(* IEC 61131-3 sources: plc-st-coding-agent/progress/evidence/f14_v3_parallel_20261112/jobs/custom_deepseek-v4pro, 102 files *)

(* ---- public-easy-01.candidate_01.st ---- *)
FUNCTION_BLOCK AutomatedFillingLineControl
VAR_INPUT
    bottleSensor : BOOL;
    cleaningConfirmButton : BOOL;
    fillingConfirmButton : BOOL;
    cappingConfirmButton : BOOL;
    packingConfirmButton : BOOL;
    finishedButton : BOOL;
END_VAR
VAR_OUTPUT
    Pump_Motor : BOOL;
    Filling_Valve : BOOL;
    Capping_Machine : BOOL;
    Packing_Machine : BOOL;
    Completion_Light : BOOL;
END_VAR
VAR
    state : INT := 0; (* 0=Idle, 1=Cleaning, 2=Filling, 3=Capping, 4=Packing, 5=Completed *)
END_VAR

CASE state OF
    0: (* Idle *)
        Pump_Motor := FALSE;
        Filling_Valve := FALSE;
        Capping_Machine := FALSE;
        Packing_Machine := FALSE;
        Completion_Light := FALSE;
        IF bottleSensor THEN
            state := 1;
        END_IF;

    1: (* Cleaning *)
        Pump_Motor := TRUE;
        Filling_Valve := FALSE;
        Capping_Machine := FALSE;
        Packing_Machine := FALSE;
        Completion_Light := FALSE;
        IF cleaningConfirmButton THEN
            state := 2;
        END_IF;

    2: (* Filling *)
        Pump_Motor := FALSE;
        Filling_Valve := TRUE;
        Capping_Machine := FALSE;
        Packing_Machine := FALSE;
        Completion_Light := FALSE;
        IF fillingConfirmButton THEN
            state := 3;
        END_IF;

    3: (* Capping *)
        Pump_Motor := FALSE;
        Filling_Valve := FALSE;
        Capping_Machine := TRUE;
        Packing_Machine := FALSE;
        Completion_Light := FALSE;
        IF cappingConfirmButton THEN
            state := 4;
        END_IF;

    4: (* Packing *)
        Pump_Motor := FALSE;
        Filling_Valve := FALSE;
        Capping_Machine := FALSE;
        Packing_Machine := TRUE;
        Completion_Light := FALSE;
        IF packingConfirmButton THEN
            state := 5;
        END_IF;

    5: (* Completed *)
        Pump_Motor := FALSE;
        Filling_Valve := FALSE;
        Capping_Machine := FALSE;
        Packing_Machine := FALSE;
        Completion_Light := TRUE;
        IF finishedButton THEN
            state := 0;
        END_IF;
END_CASE;

END_FUNCTION_BLOCK

(* ---- public-easy-01.candidate_02.st ---- *)
FUNCTION_BLOCK AutomatedFillingLineControl
VAR_INPUT
    bottleSensor : BOOL;
    cleaningConfirmButton : BOOL;
    fillingConfirmButton : BOOL;
    cappingConfirmButton : BOOL;
    packingConfirmButton : BOOL;
    finishedButton : BOOL;
END_VAR
VAR_OUTPUT
    Pump_Motor : BOOL;
    Filling_Valve : BOOL;
    Capping_Machine : BOOL;
    Packing_Machine : BOOL;
    Completion_Light : BOOL;
END_VAR
VAR
    state : INT := 0; (* 0=Idle, 1=Cleaning, 2=Filling, 3=Capping, 4=Packing, 5=Completed *)
END_VAR

CASE state OF
    0: (* Idle *)
        Pump_Motor := FALSE;
        Filling_Valve := FALSE;
        Capping_Machine := FALSE;
        Packing_Machine := FALSE;
        Completion_Light := FALSE;
        IF bottleSensor THEN
            Pump_Motor := TRUE;
            state := 1;
        END_IF;

    1: (* Cleaning *)
        Pump_Motor := TRUE;
        Filling_Valve := FALSE;
        Capping_Machine := FALSE;
        Packing_Machine := FALSE;
        Completion_Light := FALSE;
        IF cleaningConfirmButton THEN
            Pump_Motor := FALSE;
            Filling_Valve := TRUE;
            state := 2;
        END_IF;

    2: (* Filling *)
        Pump_Motor := FALSE;
        Filling_Valve := TRUE;
        Capping_Machine := FALSE;
        Packing_Machine := FALSE;
        Completion_Light := FALSE;
        IF fillingConfirmButton THEN
            Filling_Valve := FALSE;
            Capping_Machine := TRUE;
            state := 3;
        END_IF;

    3: (* Capping *)
        Pump_Motor := FALSE;
        Filling_Valve := FALSE;
        Capping_Machine := TRUE;
        Packing_Machine := FALSE;
        Completion_Light := FALSE;
        IF cappingConfirmButton THEN
            Capping_Machine := FALSE;
            Packing_Machine := TRUE;
            state := 4;
        END_IF;

    4: (* Packing *)
        Pump_Motor := FALSE;
        Filling_Valve := FALSE;
        Capping_Machine := FALSE;
        Packing_Machine := TRUE;
        Completion_Light := FALSE;
        IF packingConfirmButton THEN
            Packing_Machine := FALSE;
            Completion_Light := TRUE;
            state := 5;
        END_IF;

    5: (* Completed *)
        Pump_Motor := FALSE;
        Filling_Valve := FALSE;
        Capping_Machine := FALSE;
        Packing_Machine := FALSE;
        Completion_Light := TRUE;
        IF finishedButton THEN
            Completion_Light := FALSE;
            state := 0;
        END_IF;
END_CASE;

END_FUNCTION_BLOCK

(* ---- public-easy-01.raw_candidate_01.st ---- *)
FUNCTION_BLOCK AutomatedFillingLineControl
VAR_INPUT
    bottleSensor : BOOL;
    cleaningConfirmButton : BOOL;
    fillingConfirmButton : BOOL;
    cappingConfirmButton : BOOL;
    packingConfirmButton : BOOL;
    finishedButton : BOOL;
END_VAR
VAR_OUTPUT
    Pump_Motor : BOOL;
    Filling_Valve : BOOL;
    Capping_Machine : BOOL;
    Packing_Machine : BOOL;
    Completion_Light : BOOL;
END_VAR
VAR
    state : INT := 0; (* 0=Idle, 1=Cleaning, 2=Filling, 3=Capping, 4=Packing, 5=Completed *)
END_VAR

CASE state OF
    0: (* Idle *)
        Pump_Motor := FALSE;
        Filling_Valve := FALSE;
        Capping_Machine := FALSE;
        Packing_Machine := FALSE;
        Completion_Light := FALSE;
        IF bottleSensor THEN
            state := 1;
        END_IF;

    1: (* Cleaning *)
        Pump_Motor := TRUE;
        Filling_Valve := FALSE;
        Capping_Machine := FALSE;
        Packing_Machine := FALSE;
        Completion_Light := FALSE;
        IF cleaningConfirmButton THEN
            state := 2;
        END_IF;

    2: (* Filling *)
        Pump_Motor := FALSE;
        Filling_Valve := TRUE;
        Capping_Machine := FALSE;
        Packing_Machine := FALSE;
        Completion_Light := FALSE;
        IF fillingConfirmButton THEN
            state := 3;
        END_IF;

    3: (* Capping *)
        Pump_Motor := FALSE;
        Filling_Valve := FALSE;
        Capping_Machine := TRUE;
        Packing_Machine := FALSE;
        Completion_Light := FALSE;
        IF cappingConfirmButton THEN
            state := 4;
        END_IF;

    4: (* Packing *)
        Pump_Motor := FALSE;
        Filling_Valve := FALSE;
        Capping_Machine := FALSE;
        Packing_Machine := TRUE;
        Completion_Light := FALSE;
        IF packingConfirmButton THEN
            state := 5;
        END_IF;

    5: (* Completed *)
        Pump_Motor := FALSE;
        Filling_Valve := FALSE;
        Capping_Machine := FALSE;
        Packing_Machine := FALSE;
        Completion_Light := TRUE;
        IF finishedButton THEN
            state := 0;
        END_IF;
END_CASE;

END_FUNCTION_BLOCK

(* ---- public-easy-01.raw_candidate_02.st ---- *)
FUNCTION_BLOCK AutomatedFillingLineControl
VAR_INPUT
    bottleSensor : BOOL;
    cleaningConfirmButton : BOOL;
    fillingConfirmButton : BOOL;
    cappingConfirmButton : BOOL;
    packingConfirmButton : BOOL;
    finishedButton : BOOL;
END_VAR
VAR_OUTPUT
    Pump_Motor : BOOL;
    Filling_Valve : BOOL;
    Capping_Machine : BOOL;
    Packing_Machine : BOOL;
    Completion_Light : BOOL;
END_VAR
VAR
    state : INT := 0; (* 0=Idle, 1=Cleaning, 2=Filling, 3=Capping, 4=Packing, 5=Completed *)
END_VAR

CASE state OF
    0: (* Idle *)
        Pump_Motor := FALSE;
        Filling_Valve := FALSE;
        Capping_Machine := FALSE;
        Packing_Machine := FALSE;
        Completion_Light := FALSE;
        IF bottleSensor THEN
            Pump_Motor := TRUE;
            state := 1;
        END_IF;

    1: (* Cleaning *)
        Pump_Motor := TRUE;
        Filling_Valve := FALSE;
        Capping_Machine := FALSE;
        Packing_Machine := FALSE;
        Completion_Light := FALSE;
        IF cleaningConfirmButton THEN
            Pump_Motor := FALSE;
            Filling_Valve := TRUE;
            state := 2;
        END_IF;

    2: (* Filling *)
        Pump_Motor := FALSE;
        Filling_Valve := TRUE;
        Capping_Machine := FALSE;
        Packing_Machine := FALSE;
        Completion_Light := FALSE;
        IF fillingConfirmButton THEN
            Filling_Valve := FALSE;
            Capping_Machine := TRUE;
            state := 3;
        END_IF;

    3: (* Capping *)
        Pump_Motor := FALSE;
        Filling_Valve := FALSE;
        Capping_Machine := TRUE;
        Packing_Machine := FALSE;
        Completion_Light := FALSE;
        IF cappingConfirmButton THEN
            Capping_Machine := FALSE;
            Packing_Machine := TRUE;
            state := 4;
        END_IF;

    4: (* Packing *)
        Pump_Motor := FALSE;
        Filling_Valve := FALSE;
        Capping_Machine := FALSE;
        Packing_Machine := TRUE;
        Completion_Light := FALSE;
        IF packingConfirmButton THEN
            Packing_Machine := FALSE;
            Completion_Light := TRUE;
            state := 5;
        END_IF;

    5: (* Completed *)
        Pump_Motor := FALSE;
        Filling_Valve := FALSE;
        Capping_Machine := FALSE;
        Packing_Machine := FALSE;
        Completion_Light := TRUE;
        IF finishedButton THEN
            Completion_Light := FALSE;
            state := 0;
        END_IF;
END_CASE;

END_FUNCTION_BLOCK

(* ---- public-easy-04.candidate_01.st ---- *)
FUNCTION_BLOCK FB_JamPumpControl
VAR_INPUT
    VISCOSITY_OK : BOOL;
    PASTE_E_STOP_NC : BOOL;
    DebounceTime : TIME;
    CycleTime : TIME;
END_VAR
VAR_OUTPUT
    VFD_RUN : BOOL := FALSE;
    PUMP_MAINT_DUE : BOOL := FALSE;
    PUMP_RUNTIME_ACC : LTIME := LTIME#0s;
END_VAR
VAR
    ViscosityConditionValid : BOOL := FALSE;
    DebounceElapsed : TIME := T#0s;
    RuntimeAccumulator : LTIME := LTIME#0s;
    MaintenanceThreshold : LTIME := LTIME#500h;
END_VAR

IF NOT VISCOSITY_OK THEN
    ViscosityConditionValid := FALSE;
    DebounceElapsed := T#0s;
ELSE
    IF NOT PASTE_E_STOP_NC THEN
        DebounceElapsed := T#0s;
    ELSIF NOT ViscosityConditionValid THEN
        DebounceElapsed := DebounceElapsed + CycleTime;
        IF DebounceElapsed >= DebounceTime THEN
            ViscosityConditionValid := TRUE;
        END_IF;
    END_IF;
END_IF;

VFD_RUN := PASTE_E_STOP_NC AND ViscosityConditionValid;

IF VFD_RUN THEN
    RuntimeAccumulator := RuntimeAccumulator + TO_LTIME(CycleTime);
END_IF;

PUMP_RUNTIME_ACC := RuntimeAccumulator;
PUMP_MAINT_DUE := RuntimeAccumulator >= MaintenanceThreshold;

END_FUNCTION_BLOCK

(* ---- public-easy-04.candidate_02.st ---- *)
FUNCTION_BLOCK FB_JamPumpControl
VAR_INPUT
    VISCOSITY_OK : BOOL;
    PASTE_E_STOP_NC : BOOL;
    DebounceTime : TIME;
    CycleTime : TIME;
END_VAR
VAR_OUTPUT
    VFD_RUN : BOOL := FALSE;
    PUMP_MAINT_DUE : BOOL := FALSE;
    PUMP_RUNTIME_ACC : LTIME := LTIME#0s;
END_VAR
VAR
    ViscosityConditionValid : BOOL := FALSE;
    DebounceElapsed : TIME := T#0s;
    RuntimeAccumulator : LTIME := LTIME#0s;
    MaintenanceThreshold : LTIME := LTIME#500h;
    LastVFD_RUN : BOOL := FALSE;
END_VAR

// Debounce viscosity signal
IF NOT VISCOSITY_OK THEN
    ViscosityConditionValid := FALSE;
    DebounceElapsed := T#0s;
ELSE
    IF NOT PASTE_E_STOP_NC THEN
        // E-stop clears incomplete debounce, but keeps already valid condition
        DebounceElapsed := T#0s;
    ELSIF NOT ViscosityConditionValid THEN
        DebounceElapsed := DebounceElapsed + CycleTime;
        IF DebounceElapsed >= DebounceTime THEN
            ViscosityConditionValid := TRUE;
        END_IF;
    END_IF;
END_IF;

// VFD run permissive
VFD_RUN := PASTE_E_STOP_NC AND ViscosityConditionValid;

// Accumulate runtime, skipping the first scan after pump start
IF VFD_RUN AND NOT LastVFD_RUN THEN
    // Rising edge, do not accumulate this cycle
ELSIF VFD_RUN THEN
    RuntimeAccumulator := RuntimeAccumulator + TO_LTIME(CycleTime);
END_IF;

LastVFD_RUN := VFD_RUN;

PUMP_RUNTIME_ACC := RuntimeAccumulator;
PUMP_MAINT_DUE := RuntimeAccumulator >= MaintenanceThreshold;

END_FUNCTION_BLOCK

(* ---- public-easy-04.raw_candidate_01.st ---- *)
FUNCTION_BLOCK FB_JamPumpControl
VAR_INPUT
    VISCOSITY_OK : BOOL;
    PASTE_E_STOP_NC : BOOL;
    DebounceTime : TIME;
    CycleTime : TIME;
END_VAR
VAR_OUTPUT
    VFD_RUN : BOOL := FALSE;
    PUMP_MAINT_DUE : BOOL := FALSE;
    PUMP_RUNTIME_ACC : LTIME := LTIME#0s;
END_VAR
VAR
    ViscosityConditionValid : BOOL := FALSE;
    DebounceElapsed : TIME := T#0s;
    RuntimeAccumulator : LTIME := LTIME#0s;
    MaintenanceThreshold : LTIME := LTIME#500h;
END_VAR

IF NOT VISCOSITY_OK THEN
    ViscosityConditionValid := FALSE;
    DebounceElapsed := T#0s;
ELSE
    IF NOT PASTE_E_STOP_NC THEN
        DebounceElapsed := T#0s;
    ELSIF NOT ViscosityConditionValid THEN
        DebounceElapsed := DebounceElapsed + CycleTime;
        IF DebounceElapsed >= DebounceTime THEN
            ViscosityConditionValid := TRUE;
        END_IF;
    END_IF;
END_IF;

VFD_RUN := PASTE_E_STOP_NC AND ViscosityConditionValid;

IF VFD_RUN THEN
    RuntimeAccumulator := RuntimeAccumulator + TO_LTIME(CycleTime);
END_IF;

PUMP_RUNTIME_ACC := RuntimeAccumulator;
PUMP_MAINT_DUE := RuntimeAccumulator >= MaintenanceThreshold;

END_FUNCTION_BLOCK

(* ---- public-easy-04.raw_candidate_02.st ---- *)
FUNCTION_BLOCK FB_JamPumpControl
VAR_INPUT
    VISCOSITY_OK : BOOL;
    PASTE_E_STOP_NC : BOOL;
    DebounceTime : TIME;
    CycleTime : TIME;
END_VAR
VAR_OUTPUT
    VFD_RUN : BOOL := FALSE;
    PUMP_MAINT_DUE : BOOL := FALSE;
    PUMP_RUNTIME_ACC : LTIME := LTIME#0s;
END_VAR
VAR
    ViscosityConditionValid : BOOL := FALSE;
    DebounceElapsed : TIME := T#0s;
    RuntimeAccumulator : LTIME := LTIME#0s;
    MaintenanceThreshold : LTIME := LTIME#500h;
    LastVFD_RUN : BOOL := FALSE;
END_VAR

// Debounce viscosity signal
IF NOT VISCOSITY_OK THEN
    ViscosityConditionValid := FALSE;
    DebounceElapsed := T#0s;
ELSE
    IF NOT PASTE_E_STOP_NC THEN
        // E-stop clears incomplete debounce, but keeps already valid condition
        DebounceElapsed := T#0s;
    ELSIF NOT ViscosityConditionValid THEN
        DebounceElapsed := DebounceElapsed + CycleTime;
        IF DebounceElapsed >= DebounceTime THEN
            ViscosityConditionValid := TRUE;
        END_IF;
    END_IF;
END_IF;

// VFD run permissive
VFD_RUN := PASTE_E_STOP_NC AND ViscosityConditionValid;

// Accumulate runtime, skipping the first scan after pump start
IF VFD_RUN AND NOT LastVFD_RUN THEN
    // Rising edge, do not accumulate this cycle
ELSIF VFD_RUN THEN
    RuntimeAccumulator := RuntimeAccumulator + TO_LTIME(CycleTime);
END_IF;

LastVFD_RUN := VFD_RUN;

PUMP_RUNTIME_ACC := RuntimeAccumulator;
PUMP_MAINT_DUE := RuntimeAccumulator >= MaintenanceThreshold;

END_FUNCTION_BLOCK

(* ---- public-easy-05.candidate_01.st ---- *)
FUNCTION_BLOCK WeldGapAlarm
VAR
    TON_Init     : TON;
    TON_Debounce : TON;
    InitActive   : BOOL;
    DebounceInput: BOOL;
END_VAR

TON_Init(IN := TRUE, PT := T#5S);
InitActive := NOT TON_Init.Q;

DebounceInput := Gap_Exceeded AND NOT InitActive AND Weld_E_Stop_NC;
TON_Debounce(IN := DebounceInput, PT := DebounceTime);

Operator_Alert := TON_Debounce.Q AND Weld_E_Stop_NC AND NOT InitActive;
Weld_Soft_Start_Active := InitActive AND Weld_E_Stop_NC;

END_FUNCTION_BLOCK

(* ---- public-easy-05.candidate_02.st ---- *)
FUNCTION_BLOCK WeldGapAlarm
VAR
    Gap_Exceeded          : BOOL;  (* Input: Scanner indication that gap exceeds 1.5 mm *)
    Weld_E_Stop_NC        : BOOL;  (* Input: TRUE = emergency stop inactive; FALSE = active *)
    DebounceTime          : TIME;  (* Input: gap-signal debounce duration during normal monitoring *)

    Operator_Alert        : BOOL;  (* Output: Audible and visual alarm command *)
    Weld_Soft_Start_Active: BOOL;  (* Output: Monitoring-inhibition status during power-up init *)

    TON_Init              : TON;   (* 5-second power-up initialization timer *)
    TON_Debounce          : TON;   (* Gap-signal debounce timer *)
    InitActive            : BOOL;  (* TRUE during the 5-second initialization period *)
    DebounceInput         : BOOL;  (* Internal enable for the debounce timer *)
END_VAR

(* Power-up initialization timer: always runs for the first 5 seconds *)
TON_Init(IN := TRUE, PT := T#5S);
InitActive := NOT TON_Init.Q;

(* Debounce input is enabled only during normal monitoring (after initialization) and when E-stop is inactive *)
DebounceInput := Gap_Exceeded AND NOT InitActive AND Weld_E_Stop_NC;
TON_Debounce(IN := DebounceInput, PT := DebounceTime);

(* Operator_Alert is active when debounce has elapsed, monitoring is active, and E-stop is inactive *)
Operator_Alert := TON_Debounce.Q AND NOT InitActive AND Weld_E_Stop_NC;

(* Weld_Soft_Start_Active indicates the power-up inhibition period, but only if E-stop is inactive *)
Weld_Soft_Start_Active := InitActive AND Weld_E_Stop_NC;

END_FUNCTION_BLOCK

(* ---- public-easy-05.raw_candidate_01.st ---- *)
FUNCTION_BLOCK WeldGapAlarm
VAR
    TON_Init     : TON;
    TON_Debounce : TON;
    InitActive   : BOOL;
    DebounceInput: BOOL;
END_VAR

TON_Init(IN := TRUE, PT := T#5S);
InitActive := NOT TON_Init.Q;

DebounceInput := Gap_Exceeded AND NOT InitActive AND Weld_E_Stop_NC;
TON_Debounce(IN := DebounceInput, PT := DebounceTime);

Operator_Alert := TON_Debounce.Q AND Weld_E_Stop_NC AND NOT InitActive;
Weld_Soft_Start_Active := InitActive AND Weld_E_Stop_NC;

END_FUNCTION_BLOCK

(* ---- public-easy-05.raw_candidate_02.st ---- *)
FUNCTION_BLOCK WeldGapAlarm
VAR
    Gap_Exceeded          : BOOL;  (* Input: Scanner indication that gap exceeds 1.5 mm *)
    Weld_E_Stop_NC        : BOOL;  (* Input: TRUE = emergency stop inactive; FALSE = active *)
    DebounceTime          : TIME;  (* Input: gap-signal debounce duration during normal monitoring *)

    Operator_Alert        : BOOL;  (* Output: Audible and visual alarm command *)
    Weld_Soft_Start_Active: BOOL;  (* Output: Monitoring-inhibition status during power-up init *)

    TON_Init              : TON;   (* 5-second power-up initialization timer *)
    TON_Debounce          : TON;   (* Gap-signal debounce timer *)
    InitActive            : BOOL;  (* TRUE during the 5-second initialization period *)
    DebounceInput         : BOOL;  (* Internal enable for the debounce timer *)
END_VAR

(* Power-up initialization timer: always runs for the first 5 seconds *)
TON_Init(IN := TRUE, PT := T#5S);
InitActive := NOT TON_Init.Q;

(* Debounce input is enabled only during normal monitoring (after initialization) and when E-stop is inactive *)
DebounceInput := Gap_Exceeded AND NOT InitActive AND Weld_E_Stop_NC;
TON_Debounce(IN := DebounceInput, PT := DebounceTime);

(* Operator_Alert is active when debounce has elapsed, monitoring is active, and E-stop is inactive *)
Operator_Alert := TON_Debounce.Q AND NOT InitActive AND Weld_E_Stop_NC;

(* Weld_Soft_Start_Active indicates the power-up inhibition period, but only if E-stop is inactive *)
Weld_Soft_Start_Active := InitActive AND Weld_E_Stop_NC;

END_FUNCTION_BLOCK

(* ---- public-easy-06.candidate_01.st ---- *)
FUNCTION_BLOCK AerationBlowerDelayedStart
VAR_INPUT
    DO_LOW : BOOL;
    AERATION_E_STOP_NC : BOOL;
END_VAR
VAR_OUTPUT
    BLOWER_RUN : BOOL;
    AERATION_BLOWER_CYCLE_COUNT : UINT;
END_VAR
VAR
    startCondition : BOOL;
    runInternal : BOOL := FALSE;
    countInternal : UINT := 0;
    prevRun : BOOL := FALSE;
    fbTon : TON;
END_VAR

startCondition := DO_LOW AND AERATION_E_STOP_NC;
fbTon(IN := startCondition, PT := T#5s);
runInternal := fbTon.Q;
BLOWER_RUN := runInternal;

IF runInternal AND NOT prevRun THEN
    countInternal := countInternal + 1;
END_IF;
prevRun := runInternal;

AERATION_BLOWER_CYCLE_COUNT := countInternal;
END_FUNCTION_BLOCK

(* ---- public-easy-06.raw_candidate_01.st ---- *)
FUNCTION_BLOCK AerationBlowerDelayedStart
VAR_INPUT
    DO_LOW : BOOL;
    AERATION_E_STOP_NC : BOOL;
END_VAR
VAR_OUTPUT
    BLOWER_RUN : BOOL;
    AERATION_BLOWER_CYCLE_COUNT : UINT;
END_VAR
VAR
    startCondition : BOOL;
    runInternal : BOOL := FALSE;
    countInternal : UINT := 0;
    prevRun : BOOL := FALSE;
    fbTon : TON;
END_VAR

startCondition := DO_LOW AND AERATION_E_STOP_NC;
fbTon(IN := startCondition, PT := T#5s);
runInternal := fbTon.Q;
BLOWER_RUN := runInternal;

IF runInternal AND NOT prevRun THEN
    countInternal := countInternal + 1;
END_IF;
prevRun := runInternal;

AERATION_BLOWER_CYCLE_COUNT := countInternal;
END_FUNCTION_BLOCK

(* ---- public-hard-01.candidate_01.st ---- *)
FUNCTION_BLOCK MaterialProportioningControl
VAR CONSTANT
    STATE_IDLE : INT := 0;
    STATE_VALVE_A : INT := 1;
    STATE_VALVE_B : INT := 2;
    STATE_VALVE_C : INT := 3;
    STATE_MIXING : INT := 4;
    STATE_DONE : INT := 5;
END_VAR
VAR_INPUT
    estop : BOOL;
    opeMode : BOOL;
    valveAStart : BOOL;
    valveBStart : BOOL;
    valveCStart : BOOL;
    valveDStart : BOOL;
    mixMotorStart : BOOL;
    autoStart : BOOL;
    processMode : BOOL;
    levelSensor : INT;
    mixMotorComplete : BOOL;
END_VAR
VAR_OUTPUT
    valveARun : BOOL;
    valveBRun : BOOL;
    valveCRun : BOOL;
    valveDRun : BOOL;
    mixMotorRun : BOOL;
END_VAR
VAR
    manValveA : BOOL := FALSE;
    manValveB : BOOL := FALSE;
    manValveC : BOOL := FALSE;
    manValveD : BOOL := FALSE;
    manMixMotor : BOOL := FALSE;
    prevAutoStart : BOOL := FALSE;
    prevValveAStart : BOOL := FALSE;
    prevValveBStart : BOOL := FALSE;
    prevValveCStart : BOOL := FALSE;
    prevValveDStart : BOOL := FALSE;
    prevMixMotorStart : BOOL := FALSE;
    autoState : INT := STATE_IDLE;
END_VAR

IF NOT estop THEN
    valveARun := FALSE;
    valveBRun := FALSE;
    valveCRun := FALSE;
    valveDRun := FALSE;
    mixMotorRun := FALSE;
    manValveA := FALSE;
    manValveB := FALSE;
    manValveC := FALSE;
    manValveD := FALSE;
    manMixMotor := FALSE;
    autoState := STATE_IDLE;
ELSE
    IF NOT opeMode THEN
        IF valveAStart AND NOT prevValveAStart THEN
            manValveA := NOT manValveA;
        END_IF;
        IF valveBStart AND NOT prevValveBStart THEN
            manValveB := NOT manValveB;
        END_IF;
        IF valveCStart AND NOT prevValveCStart THEN
            manValveC := NOT manValveC;
        END_IF;
        IF valveDStart AND NOT prevValveDStart THEN
            manValveD := NOT manValveD;
        END_IF;
        IF mixMotorStart AND NOT prevMixMotorStart THEN
            manMixMotor := NOT manMixMotor;
        END_IF;
        valveARun := manValveA;
        valveBRun := manValveB;
        valveCRun := manValveC;
        valveDRun := manValveD;
        mixMotorRun := manMixMotor;
        autoState := STATE_IDLE;
    ELSE
        IF autoStart AND NOT prevAutoStart THEN
            autoState := STATE_VALVE_A;
        END_IF;
        CASE autoState OF
            STATE_IDLE:
                valveARun := FALSE;
                valveBRun := FALSE;
                valveCRun := FALSE;
                valveDRun := FALSE;
                mixMotorRun := FALSE;
            STATE_VALVE_A:
                valveARun := TRUE;
                valveBRun := FALSE;
                valveCRun := FALSE;
                valveDRun := FALSE;
                mixMotorRun := FALSE;
                IF levelSensor >= 50 THEN
                    autoState := STATE_VALVE_B;
                END_IF;
            STATE_VALVE_B:
                valveARun := FALSE;
                valveBRun := TRUE;
                valveCRun := FALSE;
                valveDRun := FALSE;
                mixMotorRun := FALSE;
                IF levelSensor >= 80 THEN
                    IF processMode THEN
                        autoState := STATE_VALVE_C;
                    ELSE
                        autoState := STATE_MIXING;
                    END_IF;
                END_IF;
            STATE_VALVE_C:
                valveARun := FALSE;
                valveBRun := FALSE;
                valveCRun := TRUE;
                valveDRun := FALSE;
                mixMotorRun := FALSE;
                IF levelSensor >= 100 THEN
                    autoState := STATE_MIXING;
                END_IF;
            STATE_MIXING:
                valveARun := FALSE;
                valveBRun := FALSE;
                valveCRun := FALSE;
                valveDRun := FALSE;
                mixMotorRun := TRUE;
                IF mixMotorComplete THEN
                    autoState := STATE_DONE;
                END_IF;
            STATE_DONE:
                valveARun := FALSE;
                valveBRun := FALSE;
                valveCRun := FALSE;
                valveDRun := TRUE;
                mixMotorRun := FALSE;
        END_CASE;
    END_IF;
END_IF;

prevAutoStart := autoStart;
prevValveAStart := valveAStart;
prevValveBStart := valveBStart;
prevValveCStart := valveCStart;
prevValveDStart := valveDStart;
prevMixMotorStart := mixMotorStart;

END_FUNCTION_BLOCK

(* ---- public-hard-01.candidate_02.st ---- *)
FUNCTION_BLOCK MaterialProportioningControl
VAR CONSTANT
    STATE_IDLE : INT := 0;
    STATE_VALVE_A : INT := 1;
    STATE_VALVE_B : INT := 2;
    STATE_VALVE_C : INT := 3;
    STATE_MIXING : INT := 4;
    STATE_DONE : INT := 5;
END_VAR
VAR_INPUT
    estop : BOOL;
    opeMode : BOOL;
    valveAStart : BOOL;
    valveBStart : BOOL;
    valveCStart : BOOL;
    valveDStart : BOOL;
    mixMotorStart : BOOL;
    autoStart : BOOL;
    processMode : BOOL;
    levelSensor : INT;
    mixMotorComplete : BOOL;
END_VAR
VAR_OUTPUT
    valveARun : BOOL;
    valveBRun : BOOL;
    valveCRun : BOOL;
    valveDRun : BOOL;
    mixMotorRun : BOOL;
END_VAR
VAR
    manValveA : BOOL := FALSE;
    manValveB : BOOL := FALSE;
    manValveC : BOOL := FALSE;
    manValveD : BOOL := FALSE;
    manMixMotor : BOOL := FALSE;
    prevAutoStart : BOOL := FALSE;
    prevValveAStart : BOOL := FALSE;
    prevValveBStart : BOOL := FALSE;
    prevValveCStart : BOOL := FALSE;
    prevValveDStart : BOOL := FALSE;
    prevMixMotorStart : BOOL := FALSE;
    autoState : INT := STATE_IDLE;
END_VAR

IF NOT estop THEN
    valveARun := FALSE;
    valveBRun := FALSE;
    valveCRun := FALSE;
    valveDRun := FALSE;
    mixMotorRun := FALSE;
    manValveA := FALSE;
    manValveB := FALSE;
    manValveC := FALSE;
    manValveD := FALSE;
    manMixMotor := FALSE;
    autoState := STATE_IDLE;
ELSE
    IF NOT opeMode THEN
        (* Manual mode *)
        IF valveAStart AND NOT prevValveAStart THEN
            manValveA := NOT manValveA;
        END_IF;
        IF valveBStart AND NOT prevValveBStart THEN
            manValveB := NOT manValveB;
        END_IF;
        IF valveCStart AND NOT prevValveCStart THEN
            manValveC := NOT manValveC;
        END_IF;
        IF valveDStart AND NOT prevValveDStart THEN
            manValveD := NOT manValveD;
        END_IF;
        IF mixMotorStart AND NOT prevMixMotorStart THEN
            manMixMotor := NOT manMixMotor;
        END_IF;
        valveARun := manValveA;
        valveBRun := manValveB;
        valveCRun := manValveC;
        valveDRun := manValveD;
        mixMotorRun := manMixMotor;
        autoState := STATE_IDLE;
    ELSE
        (* Automatic mode *)
        IF autoStart AND NOT prevAutoStart THEN
            autoState := STATE_VALVE_A;
        END_IF;

        (* State transition logic *)
        CASE autoState OF
            STATE_IDLE:
                (* No transition *)
            STATE_VALVE_A:
                IF levelSensor >= 50 THEN
                    autoState := STATE_VALVE_B;
                END_IF;
            STATE_VALVE_B:
                IF levelSensor >= 80 THEN
                    IF processMode THEN
                        autoState := STATE_VALVE_C;
                    ELSE
                        autoState := STATE_MIXING;
                    END_IF;
                END_IF;
            STATE_VALVE_C:
                IF levelSensor >= 100 THEN
                    autoState := STATE_MIXING;
                END_IF;
            STATE_MIXING:
                IF mixMotorComplete THEN
                    autoState := STATE_DONE;
                END_IF;
            STATE_DONE:
                (* Hold final state until next start *)
        END_CASE;

        (* Output based on updated state *)
        CASE autoState OF
            STATE_IDLE:
                valveARun := FALSE;
                valveBRun := FALSE;
                valveCRun := FALSE;
                valveDRun := FALSE;
                mixMotorRun := FALSE;
            STATE_VALVE_A:
                valveARun := TRUE;
                valveBRun := FALSE;
                valveCRun := FALSE;
                valveDRun := FALSE;
                mixMotorRun := FALSE;
            STATE_VALVE_B:
                valveARun := FALSE;
                valveBRun := TRUE;
                valveCRun := FALSE;
                valveDRun := FALSE;
                mixMotorRun := FALSE;
            STATE_VALVE_C:
                valveARun := FALSE;
                valveBRun := FALSE;
                valveCRun := TRUE;
                valveDRun := FALSE;
                mixMotorRun := FALSE;
            STATE_MIXING:
                valveARun := FALSE;
                valveBRun := FALSE;
                valveCRun := FALSE;
                valveDRun := FALSE;
                mixMotorRun := TRUE;
            STATE_DONE:
                valveARun := FALSE;
                valveBRun := FALSE;
                valveCRun := FALSE;
                valveDRun := TRUE;
                mixMotorRun := FALSE;
        END_CASE;
    END_IF;
END_IF;

(* Update previous input states *)
prevAutoStart := autoStart;
prevValveAStart := valveAStart;
prevValveBStart := valveBStart;
prevValveCStart := valveCStart;
prevValveDStart := valveDStart;
prevMixMotorStart := mixMotorStart;

END_FUNCTION_BLOCK

(* ---- public-hard-01.raw_candidate_01.st ---- *)
FUNCTION_BLOCK MaterialProportioningControl
VAR CONSTANT
    STATE_IDLE : INT := 0;
    STATE_VALVE_A : INT := 1;
    STATE_VALVE_B : INT := 2;
    STATE_VALVE_C : INT := 3;
    STATE_MIXING : INT := 4;
    STATE_DONE : INT := 5;
END_VAR
VAR_INPUT
    estop : BOOL;
    opeMode : BOOL;
    valveAStart : BOOL;
    valveBStart : BOOL;
    valveCStart : BOOL;
    valveDStart : BOOL;
    mixMotorStart : BOOL;
    autoStart : BOOL;
    processMode : BOOL;
    levelSensor : INT;
    mixMotorComplete : BOOL;
END_VAR
VAR_OUTPUT
    valveARun : BOOL;
    valveBRun : BOOL;
    valveCRun : BOOL;
    valveDRun : BOOL;
    mixMotorRun : BOOL;
END_VAR
VAR
    manValveA : BOOL := FALSE;
    manValveB : BOOL := FALSE;
    manValveC : BOOL := FALSE;
    manValveD : BOOL := FALSE;
    manMixMotor : BOOL := FALSE;
    prevAutoStart : BOOL := FALSE;
    prevValveAStart : BOOL := FALSE;
    prevValveBStart : BOOL := FALSE;
    prevValveCStart : BOOL := FALSE;
    prevValveDStart : BOOL := FALSE;
    prevMixMotorStart : BOOL := FALSE;
    autoState : INT := STATE_IDLE;
END_VAR

IF NOT estop THEN
    valveARun := FALSE;
    valveBRun := FALSE;
    valveCRun := FALSE;
    valveDRun := FALSE;
    mixMotorRun := FALSE;
    manValveA := FALSE;
    manValveB := FALSE;
    manValveC := FALSE;
    manValveD := FALSE;
    manMixMotor := FALSE;
    autoState := STATE_IDLE;
ELSE
    IF NOT opeMode THEN
        IF valveAStart AND NOT prevValveAStart THEN
            manValveA := NOT manValveA;
        END_IF;
        IF valveBStart AND NOT prevValveBStart THEN
            manValveB := NOT manValveB;
        END_IF;
        IF valveCStart AND NOT prevValveCStart THEN
            manValveC := NOT manValveC;
        END_IF;
        IF valveDStart AND NOT prevValveDStart THEN
            manValveD := NOT manValveD;
        END_IF;
        IF mixMotorStart AND NOT prevMixMotorStart THEN
            manMixMotor := NOT manMixMotor;
        END_IF;
        valveARun := manValveA;
        valveBRun := manValveB;
        valveCRun := manValveC;
        valveDRun := manValveD;
        mixMotorRun := manMixMotor;
        autoState := STATE_IDLE;
    ELSE
        IF autoStart AND NOT prevAutoStart THEN
            autoState := STATE_VALVE_A;
        END_IF;
        CASE autoState OF
            STATE_IDLE:
                valveARun := FALSE;
                valveBRun := FALSE;
                valveCRun := FALSE;
                valveDRun := FALSE;
                mixMotorRun := FALSE;
            STATE_VALVE_A:
                valveARun := TRUE;
                valveBRun := FALSE;
                valveCRun := FALSE;
                valveDRun := FALSE;
                mixMotorRun := FALSE;
                IF levelSensor >= 50 THEN
                    autoState := STATE_VALVE_B;
                END_IF;
            STATE_VALVE_B:
                valveARun := FALSE;
                valveBRun := TRUE;
                valveCRun := FALSE;
                valveDRun := FALSE;
                mixMotorRun := FALSE;
                IF levelSensor >= 80 THEN
                    IF processMode THEN
                        autoState := STATE_VALVE_C;
                    ELSE
                        autoState := STATE_MIXING;
                    END_IF;
                END_IF;
            STATE_VALVE_C:
                valveARun := FALSE;
                valveBRun := FALSE;
                valveCRun := TRUE;
                valveDRun := FALSE;
                mixMotorRun := FALSE;
                IF levelSensor >= 100 THEN
                    autoState := STATE_MIXING;
                END_IF;
            STATE_MIXING:
                valveARun := FALSE;
                valveBRun := FALSE;
                valveCRun := FALSE;
                valveDRun := FALSE;
                mixMotorRun := TRUE;
                IF mixMotorComplete THEN
                    autoState := STATE_DONE;
                END_IF;
            STATE_DONE:
                valveARun := FALSE;
                valveBRun := FALSE;
                valveCRun := FALSE;
                valveDRun := TRUE;
                mixMotorRun := FALSE;
        END_CASE;
    END_IF;
END_IF;

prevAutoStart := autoStart;
prevValveAStart := valveAStart;
prevValveBStart := valveBStart;
prevValveCStart := valveCStart;
prevValveDStart := valveDStart;
prevMixMotorStart := mixMotorStart;

END_FUNCTION_BLOCK

(* ---- public-hard-01.raw_candidate_02.st ---- *)
FUNCTION_BLOCK MaterialProportioningControl
VAR CONSTANT
    STATE_IDLE : INT := 0;
    STATE_VALVE_A : INT := 1;
    STATE_VALVE_B : INT := 2;
    STATE_VALVE_C : INT := 3;
    STATE_MIXING : INT := 4;
    STATE_DONE : INT := 5;
END_VAR
VAR_INPUT
    estop : BOOL;
    opeMode : BOOL;
    valveAStart : BOOL;
    valveBStart : BOOL;
    valveCStart : BOOL;
    valveDStart : BOOL;
    mixMotorStart : BOOL;
    autoStart : BOOL;
    processMode : BOOL;
    levelSensor : INT;
    mixMotorComplete : BOOL;
END_VAR
VAR_OUTPUT
    valveARun : BOOL;
    valveBRun : BOOL;
    valveCRun : BOOL;
    valveDRun : BOOL;
    mixMotorRun : BOOL;
END_VAR
VAR
    manValveA : BOOL := FALSE;
    manValveB : BOOL := FALSE;
    manValveC : BOOL := FALSE;
    manValveD : BOOL := FALSE;
    manMixMotor : BOOL := FALSE;
    prevAutoStart : BOOL := FALSE;
    prevValveAStart : BOOL := FALSE;
    prevValveBStart : BOOL := FALSE;
    prevValveCStart : BOOL := FALSE;
    prevValveDStart : BOOL := FALSE;
    prevMixMotorStart : BOOL := FALSE;
    autoState : INT := STATE_IDLE;
END_VAR

IF NOT estop THEN
    valveARun := FALSE;
    valveBRun := FALSE;
    valveCRun := FALSE;
    valveDRun := FALSE;
    mixMotorRun := FALSE;
    manValveA := FALSE;
    manValveB := FALSE;
    manValveC := FALSE;
    manValveD := FALSE;
    manMixMotor := FALSE;
    autoState := STATE_IDLE;
ELSE
    IF NOT opeMode THEN
        (* Manual mode *)
        IF valveAStart AND NOT prevValveAStart THEN
            manValveA := NOT manValveA;
        END_IF;
        IF valveBStart AND NOT prevValveBStart THEN
            manValveB := NOT manValveB;
        END_IF;
        IF valveCStart AND NOT prevValveCStart THEN
            manValveC := NOT manValveC;
        END_IF;
        IF valveDStart AND NOT prevValveDStart THEN
            manValveD := NOT manValveD;
        END_IF;
        IF mixMotorStart AND NOT prevMixMotorStart THEN
            manMixMotor := NOT manMixMotor;
        END_IF;
        valveARun := manValveA;
        valveBRun := manValveB;
        valveCRun := manValveC;
        valveDRun := manValveD;
        mixMotorRun := manMixMotor;
        autoState := STATE_IDLE;
    ELSE
        (* Automatic mode *)
        IF autoStart AND NOT prevAutoStart THEN
            autoState := STATE_VALVE_A;
        END_IF;

        (* State transition logic *)
        CASE autoState OF
            STATE_IDLE:
                (* No transition *)
            STATE_VALVE_A:
                IF levelSensor >= 50 THEN
                    autoState := STATE_VALVE_B;
                END_IF;
            STATE_VALVE_B:
                IF levelSensor >= 80 THEN
                    IF processMode THEN
                        autoState := STATE_VALVE_C;
                    ELSE
                        autoState := STATE_MIXING;
                    END_IF;
                END_IF;
            STATE_VALVE_C:
                IF levelSensor >= 100 THEN
                    autoState := STATE_MIXING;
                END_IF;
            STATE_MIXING:
                IF mixMotorComplete THEN
                    autoState := STATE_DONE;
                END_IF;
            STATE_DONE:
                (* Hold final state until next start *)
        END_CASE;

        (* Output based on updated state *)
        CASE autoState OF
            STATE_IDLE:
                valveARun := FALSE;
                valveBRun := FALSE;
                valveCRun := FALSE;
                valveDRun := FALSE;
                mixMotorRun := FALSE;
            STATE_VALVE_A:
                valveARun := TRUE;
                valveBRun := FALSE;
                valveCRun := FALSE;
                valveDRun := FALSE;
                mixMotorRun := FALSE;
            STATE_VALVE_B:
                valveARun := FALSE;
                valveBRun := TRUE;
                valveCRun := FALSE;
                valveDRun := FALSE;
                mixMotorRun := FALSE;
            STATE_VALVE_C:
                valveARun := FALSE;
                valveBRun := FALSE;
                valveCRun := TRUE;
                valveDRun := FALSE;
                mixMotorRun := FALSE;
            STATE_MIXING:
                valveARun := FALSE;
                valveBRun := FALSE;
                valveCRun := FALSE;
                valveDRun := FALSE;
                mixMotorRun := TRUE;
            STATE_DONE:
                valveARun := FALSE;
                valveBRun := FALSE;
                valveCRun := FALSE;
                valveDRun := TRUE;
                mixMotorRun := FALSE;
        END_CASE;
    END_IF;
END_IF;

(* Update previous input states *)
prevAutoStart := autoStart;
prevValveAStart := valveAStart;
prevValveBStart := valveBStart;
prevValveCStart := valveCStart;
prevValveDStart := valveDStart;
prevMixMotorStart := mixMotorStart;

END_FUNCTION_BLOCK

(* ---- public-hard-02.candidate_01.st ---- *)
FUNCTION_BLOCK FlexibleProcessingControl
VAR_INPUT
    processLength : USINT;
    sensor1 : BOOL;
    sensor2 : BOOL;
    sensor3 : BOOL;
    sensor4 : BOOL;
    sensor5 : BOOL;
    station1Start : BOOL;
    station2Complete : BOOL;
    station3Complete : BOOL;
    station4Complete : BOOL;
    processSequence : ARRAY[1..8] OF USINT;
END_VAR
VAR_OUTPUT
    conveyorLeft : BOOL;
    conveyorRight : BOOL;
END_VAR
VAR
    state : USINT := 0; (* 0: Idle, 1: Moving, 2: Processing *)
    seqIndex : USINT := 1;
    currentStation : USINT := 1;
    moveTarget : USINT := 1;

    lastStart : BOOL := FALSE;
    lastComp2 : BOOL := FALSE;
    lastComp3 : BOOL := FALSE;
    lastComp4 : BOOL := FALSE;

    startRise : BOOL := FALSE;
    comp2Rise : BOOL := FALSE;
    comp3Rise : BOOL := FALSE;
    comp4Rise : BOOL := FALSE;

    arrived : BOOL := FALSE;
    completion : BOOL := FALSE;
END_VAR

(* Input edge detection *)
startRise := station1Start AND NOT lastStart;
lastStart := station1Start;

comp2Rise := station2Complete AND NOT lastComp2;
lastComp2 := station2Complete;

comp3Rise := station3Complete AND NOT lastComp3;
lastComp3 := station3Complete;

comp4Rise := station4Complete AND NOT lastComp4;
lastComp4 := station4Complete;

(* Default outputs *)
conveyorLeft := FALSE;
conveyorRight := FALSE;

CASE state OF
    0: (* Idle *)
        IF sensor1 AND startRise THEN
            IF processLength >= 1 THEN
                seqIndex := 1;
                currentStation := 1;
                moveTarget := processSequence[1];
                state := 1;
            END_IF;
        END_IF;

    1: (* Moving *)
        IF moveTarget > currentStation THEN
            conveyorRight := TRUE;
            conveyorLeft := FALSE;
        ELSIF moveTarget < currentStation THEN
            conveyorLeft := TRUE;
            conveyorRight := FALSE;
        ELSE
            conveyorLeft := FALSE;
            conveyorRight := FALSE;
        END_IF;

        CASE moveTarget OF
            1: arrived := sensor1;
            2: arrived := sensor2;
            3: arrived := sensor3;
            4: arrived := sensor4;
            5: arrived := sensor5;
        ELSE
            arrived := FALSE;
        END_CASE;

        IF arrived THEN
            conveyorLeft := FALSE;
            conveyorRight := FALSE;
            currentStation := moveTarget;

            IF moveTarget = 5 THEN
                state := 0; (* Finished: delivered to output station *)
            ELSE
                state := 2; (* Wait for processing completion *)
            END_IF;
        END_IF;

    2: (* Processing *)
        conveyorLeft := FALSE;
        conveyorRight := FALSE;

        CASE currentStation OF
            2: completion := comp2Rise;
            3: completion := comp3Rise;
            4: completion := comp4Rise;
        ELSE
            completion := FALSE;
        END_CASE;

        IF completion THEN
            IF seqIndex < processLength THEN
                seqIndex := seqIndex + 1;
                moveTarget := processSequence[seqIndex];

                IF moveTarget = currentStation THEN
                    state := 2; (* Same station: wait for next completion *)
                ELSE
                    state := 1; (* Move to next station *)
                END_IF;
            ELSE
                state := 0; (* Safety: no further sequence entry available *)
            END_IF;
        END_IF;
END_CASE;

END_FUNCTION_BLOCK

(* ---- public-hard-02.raw_candidate_01.st ---- *)
FUNCTION_BLOCK FlexibleProcessingControl
VAR_INPUT
    processLength : USINT;
    sensor1 : BOOL;
    sensor2 : BOOL;
    sensor3 : BOOL;
    sensor4 : BOOL;
    sensor5 : BOOL;
    station1Start : BOOL;
    station2Complete : BOOL;
    station3Complete : BOOL;
    station4Complete : BOOL;
    processSequence : ARRAY[1..8] OF USINT;
END_VAR
VAR_OUTPUT
    conveyorLeft : BOOL;
    conveyorRight : BOOL;
END_VAR
VAR
    state : USINT := 0; (* 0: Idle, 1: Moving, 2: Processing *)
    seqIndex : USINT := 1;
    currentStation : USINT := 1;
    moveTarget : USINT := 1;

    lastStart : BOOL := FALSE;
    lastComp2 : BOOL := FALSE;
    lastComp3 : BOOL := FALSE;
    lastComp4 : BOOL := FALSE;

    startRise : BOOL := FALSE;
    comp2Rise : BOOL := FALSE;
    comp3Rise : BOOL := FALSE;
    comp4Rise : BOOL := FALSE;

    arrived : BOOL := FALSE;
    completion : BOOL := FALSE;
END_VAR

(* Input edge detection *)
startRise := station1Start AND NOT lastStart;
lastStart := station1Start;

comp2Rise := station2Complete AND NOT lastComp2;
lastComp2 := station2Complete;

comp3Rise := station3Complete AND NOT lastComp3;
lastComp3 := station3Complete;

comp4Rise := station4Complete AND NOT lastComp4;
lastComp4 := station4Complete;

(* Default outputs *)
conveyorLeft := FALSE;
conveyorRight := FALSE;

CASE state OF
    0: (* Idle *)
        IF sensor1 AND startRise THEN
            IF processLength >= 1 THEN
                seqIndex := 1;
                currentStation := 1;
                moveTarget := processSequence[1];
                state := 1;
            END_IF
        END_IF

    1: (* Moving *)
        IF moveTarget > currentStation THEN
            conveyorRight := TRUE;
            conveyorLeft := FALSE;
        ELSIF moveTarget < currentStation THEN
            conveyorLeft := TRUE;
            conveyorRight := FALSE;
        ELSE
            conveyorLeft := FALSE;
            conveyorRight := FALSE;
        END_IF

        CASE moveTarget OF
            1: arrived := sensor1;
            2: arrived := sensor2;
            3: arrived := sensor3;
            4: arrived := sensor4;
            5: arrived := sensor5;
        ELSE
            arrived := FALSE;
        END_CASE

        IF arrived THEN
            conveyorLeft := FALSE;
            conveyorRight := FALSE;
            currentStation := moveTarget;

            IF moveTarget = 5 THEN
                state := 0; (* Finished: delivered to output station *)
            ELSE
                state := 2; (* Wait for processing completion *)
            END_IF
        END_IF

    2: (* Processing *)
        conveyorLeft := FALSE;
        conveyorRight := FALSE;

        CASE currentStation OF
            2: completion := comp2Rise;
            3: completion := comp3Rise;
            4: completion := comp4Rise;
        ELSE
            completion := FALSE;
        END_CASE

        IF completion THEN
            IF seqIndex < processLength THEN
                seqIndex := seqIndex + 1;
                moveTarget := processSequence[seqIndex];

                IF moveTarget = currentStation THEN
                    state := 2; (* Same station: wait for next completion *)
                ELSE
                    state := 1; (* Move to next station *)
                END_IF
            ELSE
                state := 0; (* Safety: no further sequence entry available *)
            END_IF
        END_IF
END_CASE

END_FUNCTION_BLOCK

(* ---- public-hard-03.candidate_01.st ---- *)
TYPE ST_Recipe :
STRUCT
    recipeID : INT;
    ingredientType : INT;
    ingredientRatio : REAL;
    productionTemperature : REAL;
END_STRUCT;
END_TYPE;

FUNCTION_BLOCK RecipeManagement
VAR_INPUT
    addRecipe : BOOL;
    deleteRecipe : BOOL;
    modifyRecipe : BOOL;
    queryRecipe : BOOL;
    recipeIn : ST_Recipe;
END_VAR
VAR_OUTPUT
    recipeAdded : BOOL;
    recipeDeleted : BOOL;
    recipeModified : BOOL;
    recipeQueryResult : ST_Recipe;
    error : BOOL;
    status : WORD;
END_VAR
VAR_IN_OUT
    recipe : ARRAY[1..10] OF ST_Recipe;
END_VAR
VAR
    i : INT;
    foundIndex : INT;
    emptyIndex : INT;
    duplicate : BOOL;
END_VAR

    recipeAdded := FALSE;
    recipeDeleted := FALSE;
    recipeModified := FALSE;
    error := FALSE;
    status := 0;
    recipeQueryResult.recipeID := 0;
    recipeQueryResult.ingredientType := 0;
    recipeQueryResult.ingredientRatio := 0.0;
    recipeQueryResult.productionTemperature := 0.0;
    duplicate := FALSE;
    foundIndex := 0;
    emptyIndex := 0;

    IF addRecipe THEN
        duplicate := FALSE;
        foundIndex := 0;
        FOR i := 1 TO 10 DO
            IF recipe[i].recipeID <> 0 AND recipe[i].recipeID = recipeIn.recipeID THEN
                duplicate := TRUE;
                foundIndex := i;
                EXIT;
            END_IF;
        END_FOR;

        IF duplicate THEN
            error := TRUE;
            status := 16#8002;
        ELSE
            emptyIndex := 0;
            FOR i := 1 TO 10 DO
                IF recipe[i].recipeID = 0 THEN
                    emptyIndex := i;
                    EXIT;
                END_IF;
            END_FOR;
            IF emptyIndex = 0 THEN
                error := TRUE;
                status := 16#8003;
            ELSE
                recipe[emptyIndex] := recipeIn;
                recipeAdded := TRUE;
            END_IF;
        END_IF;

    ELSIF deleteRecipe THEN
        foundIndex := 0;
        FOR i := 1 TO 10 DO
            IF recipe[i].recipeID <> 0 AND recipe[i].recipeID = recipeIn.recipeID THEN
                foundIndex := i;
                EXIT;
            END_IF;
        END_FOR;
        IF foundIndex = 0 THEN
            error := TRUE;
            status := 16#8004;
        ELSE
            recipe[foundIndex].recipeID := 0;
            recipe[foundIndex].ingredientType := 0;
            recipe[foundIndex].ingredientRatio := 0.0;
            recipe[foundIndex].productionTemperature := 0.0;
            recipeDeleted := TRUE;
        END_IF;

    ELSIF modifyRecipe THEN
        foundIndex := 0;
        FOR i := 1 TO 10 DO
            IF recipe[i].recipeID <> 0 AND recipe[i].recipeID = recipeIn.recipeID THEN
                foundIndex := i;
                EXIT;
            END_IF;
        END_FOR;
        IF foundIndex = 0 THEN
            error := TRUE;
            status := 16#8005;
        ELSE
            recipe[foundIndex] := recipeIn;
            recipeModified := TRUE;
        END_IF;

    ELSIF queryRecipe THEN
        foundIndex := 0;
        FOR i := 1 TO 10 DO
            IF recipe[i].recipeID <> 0 AND recipe[i].recipeID = recipeIn.recipeID THEN
                foundIndex := i;
                EXIT;
            END_IF;
        END_FOR;
        IF foundIndex = 0 THEN
            error := TRUE;
            status := 16#8001;
        ELSE
            recipeQueryResult := recipe[foundIndex];
        END_IF;
    END_IF;

END_FUNCTION_BLOCK

(* ---- public-hard-03.candidate_02.st ---- *)
TYPE ST_Recipe :
STRUCT
    recipeID : INT;
    ingredientType : INT;
    ingredientRatio : REAL;
    productionTemperature : REAL;
END_STRUCT;
END_TYPE;

FUNCTION_BLOCK RecipeManagement
VAR_INPUT
    addRecipe : BOOL;
    deleteRecipe : BOOL;
    modifyRecipe : BOOL;
    queryRecipe : BOOL;
    recipeIn : ST_Recipe;
END_VAR
VAR_OUTPUT
    recipeAdded : BOOL;
    recipeDeleted : BOOL;
    recipeModified : BOOL;
    recipeQueryResult : ST_Recipe;
    error : BOOL;
    status : WORD;
END_VAR
VAR_IN_OUT
    recipe : ARRAY[1..10] OF ST_Recipe;
END_VAR
VAR
    i : INT;
    foundIndex : INT;
    emptyIndex : INT;
    duplicate : BOOL;
END_VAR

    recipeAdded := FALSE;
    recipeDeleted := FALSE;
    recipeModified := FALSE;
    error := FALSE;
    status := 0;
    recipeQueryResult.recipeID := 0;
    recipeQueryResult.ingredientType := 0;
    recipeQueryResult.ingredientRatio := 0.0;
    recipeQueryResult.productionTemperature := 0.0;
    duplicate := FALSE;
    foundIndex := 0;
    emptyIndex := 0;

    IF addRecipe THEN
        duplicate := FALSE;
        foundIndex := 0;
        FOR i := 1 TO 10 DO
            IF recipe[i].recipeID <> 0 AND recipe[i].recipeID = recipeIn.recipeID THEN
                duplicate := TRUE;
                foundIndex := i;
                EXIT;
            END_IF;
        END_FOR;

        IF duplicate THEN
            error := TRUE;
            status := 16#8002;
        ELSE
            emptyIndex := 0;
            FOR i := 1 TO 10 DO
                IF recipe[i].recipeID = 0 THEN
                    emptyIndex := i;
                    EXIT;
                END_IF;
            END_FOR;
            IF emptyIndex = 0 THEN
                error := TRUE;
                status := 16#8003;
            ELSE
                recipe[emptyIndex] := recipeIn;
                recipeAdded := TRUE;
            END_IF;
        END_IF;

    ELSIF deleteRecipe THEN
        foundIndex := 0;
        FOR i := 1 TO 10 DO
            IF recipe[i].recipeID <> 0 AND recipe[i].recipeID = recipeIn.recipeID THEN
                foundIndex := i;
                EXIT;
            END_IF;
        END_FOR;
        IF foundIndex = 0 THEN
            error := TRUE;
            status := 16#8004;
        ELSE
            recipe[foundIndex].recipeID := 0;
            recipe[foundIndex].ingredientType := 0;
            recipe[foundIndex].ingredientRatio := 0.0;
            recipe[foundIndex].productionTemperature := 0.0;
            recipeDeleted := TRUE;
        END_IF;

    ELSIF modifyRecipe THEN
        foundIndex := 0;
        FOR i := 1 TO 10 DO
            IF recipe[i].recipeID <> 0 AND recipe[i].recipeID = recipeIn.recipeID THEN
                foundIndex := i;
                EXIT;
            END_IF;
        END_FOR;
        IF foundIndex = 0 THEN
            error := TRUE;
            status := 16#8005;
        ELSE
            recipe[foundIndex] := recipeIn;
            recipeModified := TRUE;
        END_IF;

    ELSIF queryRecipe THEN
        foundIndex := 0;
        FOR i := 1 TO 10 DO
            IF recipe[i].recipeID <> 0 AND recipe[i].recipeID = recipeIn.recipeID THEN
                foundIndex := i;
                EXIT;
            END_IF;
        END_FOR;
        IF foundIndex = 0 THEN
            error := TRUE;
            status := 16#8001;
        ELSE
            recipeQueryResult := recipe[foundIndex];
        END_IF;
    END_IF;

END_FUNCTION_BLOCK

(* ---- public-hard-03.raw_candidate_01.st ---- *)
TYPE ST_Recipe :
STRUCT
    recipeID : INT;
    ingredientType : INT;
    ingredientRatio : REAL;
    productionTemperature : REAL;
END_STRUCT
END_TYPE

FUNCTION_BLOCK RecipeManagement
VAR_INPUT
    addRecipe : BOOL;
    deleteRecipe : BOOL;
    modifyRecipe : BOOL;
    queryRecipe : BOOL;
    recipeIn : ST_Recipe;
END_VAR
VAR_OUTPUT
    recipeAdded : BOOL;
    recipeDeleted : BOOL;
    recipeModified : BOOL;
    recipeQueryResult : ST_Recipe;
    error : BOOL;
    status : WORD;
END_VAR
VAR_IN_OUT
    recipe : ARRAY[1..10] OF ST_Recipe;
END_VAR
VAR
    i : INT;
    foundIndex : INT;
    emptyIndex : INT;
    duplicate : BOOL;
END_VAR

    recipeAdded := FALSE;
    recipeDeleted := FALSE;
    recipeModified := FALSE;
    error := FALSE;
    status := 0;
    recipeQueryResult.recipeID := 0;
    recipeQueryResult.ingredientType := 0;
    recipeQueryResult.ingredientRatio := 0.0;
    recipeQueryResult.productionTemperature := 0.0;
    duplicate := FALSE;
    foundIndex := 0;
    emptyIndex := 0;

    IF addRecipe THEN
        duplicate := FALSE;
        foundIndex := 0;
        FOR i := 1 TO 10 DO
            IF recipe[i].recipeID <> 0 AND recipe[i].recipeID = recipeIn.recipeID THEN
                duplicate := TRUE;
                foundIndex := i;
                EXIT;
            END_IF;
        END_FOR;

        IF duplicate THEN
            error := TRUE;
            status := 16#8002;
        ELSE
            emptyIndex := 0;
            FOR i := 1 TO 10 DO
                IF recipe[i].recipeID = 0 THEN
                    emptyIndex := i;
                    EXIT;
                END_IF;
            END_FOR;
            IF emptyIndex = 0 THEN
                error := TRUE;
                status := 16#8003;
            ELSE
                recipe[emptyIndex] := recipeIn;
                recipeAdded := TRUE;
            END_IF;
        END_IF;

    ELSIF deleteRecipe THEN
        foundIndex := 0;
        FOR i := 1 TO 10 DO
            IF recipe[i].recipeID <> 0 AND recipe[i].recipeID = recipeIn.recipeID THEN
                foundIndex := i;
                EXIT;
            END_IF;
        END_FOR;
        IF foundIndex = 0 THEN
            error := TRUE;
            status := 16#8004;
        ELSE
            recipe[foundIndex].recipeID := 0;
            recipe[foundIndex].ingredientType := 0;
            recipe[foundIndex].ingredientRatio := 0.0;
            recipe[foundIndex].productionTemperature := 0.0;
            recipeDeleted := TRUE;
        END_IF;

    ELSIF modifyRecipe THEN
        foundIndex := 0;
        FOR i := 1 TO 10 DO
            IF recipe[i].recipeID <> 0 AND recipe[i].recipeID = recipeIn.recipeID THEN
                foundIndex := i;
                EXIT;
            END_IF;
        END_FOR;
        IF foundIndex = 0 THEN
            error := TRUE;
            status := 16#8005;
        ELSE
            recipe[foundIndex] := recipeIn;
            recipeModified := TRUE;
        END_IF;

    ELSIF queryRecipe THEN
        foundIndex := 0;
        FOR i := 1 TO 10 DO
            IF recipe[i].recipeID <> 0 AND recipe[i].recipeID = recipeIn.recipeID THEN
                foundIndex := i;
                EXIT;
            END_IF;
        END_FOR;
        IF foundIndex = 0 THEN
            error := TRUE;
            status := 16#8001;
        ELSE
            recipeQueryResult := recipe[foundIndex];
        END_IF;
    END_IF;

END_FUNCTION_BLOCK

(* ---- public-hard-03.raw_candidate_02.st ---- *)
TYPE ST_Recipe :
STRUCT
    recipeID : INT;
    ingredientType : INT;
    ingredientRatio : REAL;
    productionTemperature : REAL;
END_STRUCT
END_TYPE

FUNCTION_BLOCK RecipeManagement
VAR_INPUT
    addRecipe : BOOL;
    deleteRecipe : BOOL;
    modifyRecipe : BOOL;
    queryRecipe : BOOL;
    recipeIn : ST_Recipe;
END_VAR
VAR_OUTPUT
    recipeAdded : BOOL;
    recipeDeleted : BOOL;
    recipeModified : BOOL;
    recipeQueryResult : ST_Recipe;
    error : BOOL;
    status : WORD;
END_VAR
VAR_IN_OUT
    recipe : ARRAY[1..10] OF ST_Recipe;
END_VAR
VAR
    i : INT;
    foundIndex : INT;
    emptyIndex : INT;
    duplicate : BOOL;
END_VAR

    recipeAdded := FALSE;
    recipeDeleted := FALSE;
    recipeModified := FALSE;
    error := FALSE;
    status := 0;
    recipeQueryResult.recipeID := 0;
    recipeQueryResult.ingredientType := 0;
    recipeQueryResult.ingredientRatio := 0.0;
    recipeQueryResult.productionTemperature := 0.0;
    duplicate := FALSE;
    foundIndex := 0;
    emptyIndex := 0;

    IF addRecipe THEN
        duplicate := FALSE;
        foundIndex := 0;
        FOR i := 1 TO 10 DO
            IF recipe[i].recipeID <> 0 AND recipe[i].recipeID = recipeIn.recipeID THEN
                duplicate := TRUE;
                foundIndex := i;
                EXIT;
            END_IF;
        END_FOR;

        IF duplicate THEN
            error := TRUE;
            status := 16#8002;
        ELSE
            emptyIndex := 0;
            FOR i := 1 TO 10 DO
                IF recipe[i].recipeID = 0 THEN
                    emptyIndex := i;
                    EXIT;
                END_IF;
            END_FOR;
            IF emptyIndex = 0 THEN
                error := TRUE;
                status := 16#8003;
            ELSE
                recipe[emptyIndex] := recipeIn;
                recipeAdded := TRUE;
            END_IF;
        END_IF;

    ELSIF deleteRecipe THEN
        foundIndex := 0;
        FOR i := 1 TO 10 DO
            IF recipe[i].recipeID <> 0 AND recipe[i].recipeID = recipeIn.recipeID THEN
                foundIndex := i;
                EXIT;
            END_IF;
        END_FOR;
        IF foundIndex = 0 THEN
            error := TRUE;
            status := 16#8004;
        ELSE
            recipe[foundIndex].recipeID := 0;
            recipe[foundIndex].ingredientType := 0;
            recipe[foundIndex].ingredientRatio := 0.0;
            recipe[foundIndex].productionTemperature := 0.0;
            recipeDeleted := TRUE;
        END_IF;

    ELSIF modifyRecipe THEN
        foundIndex := 0;
        FOR i := 1 TO 10 DO
            IF recipe[i].recipeID <> 0 AND recipe[i].recipeID = recipeIn.recipeID THEN
                foundIndex := i;
                EXIT;
            END_IF;
        END_FOR;
        IF foundIndex = 0 THEN
            error := TRUE;
            status := 16#8005;
        ELSE
            recipe[foundIndex] := recipeIn;
            recipeModified := TRUE;
        END_IF;

    ELSIF queryRecipe THEN
        foundIndex := 0;
        FOR i := 1 TO 10 DO
            IF recipe[i].recipeID <> 0 AND recipe[i].recipeID = recipeIn.recipeID THEN
                foundIndex := i;
                EXIT;
            END_IF;
        END_FOR;
        IF foundIndex = 0 THEN
            error := TRUE;
            status := 16#8001;
        ELSE
            recipeQueryResult := recipe[foundIndex];
        END_IF;
    END_IF;

END_FUNCTION_BLOCK

(* ---- public-hard-04.candidate_01.st ---- *)
FUNCTION_BLOCK FB
VAR_INPUT
    enqueue : BOOL;
    dequeue : BOOL;
    reset : BOOL;
END_VAR
VAR_OUTPUT
    elementCount : DINT;
    status : WORD;
END_VAR
VAR_IN_OUT
    item : VARIANT;
    buffer : VARIANT;
END_VAR
VAR
    head : DINT := 0;
    tail : DINT := 0;
    count : DINT := 0;
    capacity : DINT := 0;
    elemSize : DINT := 0;
    initialized : BOOL := FALSE;
    prevEnqueue : BOOL := FALSE;
    prevDequeue : BOOL := FALSE;
    enqEdge : BOOL;
    deqEdge : BOOL;
    bufferAddr : PVOID;
    itemAddr : PVOID;
    bufferSize : DINT;
    itemSize : DINT;
    destAddr : PVOID;
    srcAddr : PVOID;
    copyLen : UDINT;
END_VAR

status := 16#0000;

IF NOT initialized THEN
    bufferSize := __VARINFO(buffer).diSize;
    itemSize := __VARINFO(item).diSize;
    IF (bufferSize > 0) AND (itemSize > 0) THEN
        elemSize := itemSize;
        capacity := bufferSize / elemSize;
        bufferAddr := __VARINFO(buffer).pvAddress;
        itemAddr := __VARINFO(item).pvAddress;
        head := 0;
        tail := 0;
        count := 0;
        initialized := TRUE;
    ELSE
        elementCount := 0;
        RETURN;
    END_IF;
END_IF;

enqEdge := enqueue AND NOT prevEnqueue;
deqEdge := dequeue AND NOT prevDequeue;
prevEnqueue := enqueue;
prevDequeue := dequeue;

IF reset THEN
    head := 0;
    tail := 0;
    count := 0;
    elementCount := 0;
    status := 16#0000;
    RETURN;
END_IF;

IF enqEdge THEN
    IF count >= capacity THEN
        status := 16#8002;
    ELSE
        destAddr := bufferAddr + (tail * elemSize);
        srcAddr := itemAddr;
        copyLen := TO_UDINT(elemSize);
        SysMemCpy(destAddr, srcAddr, copyLen);
        tail := tail + 1;
        IF tail >= capacity THEN
            tail := 0;
        END_IF;
        count := count + 1;
        status := 16#0000;
    END_IF;
END_IF;

IF deqEdge THEN
    IF count = 0 THEN
        status := 16#8001;
    ELSE
        srcAddr := bufferAddr + (head * elemSize);
        destAddr := itemAddr;
        copyLen := TO_UDINT(elemSize);
        SysMemCpy(destAddr, srcAddr, copyLen);
        head := head + 1;
        IF head >= capacity THEN
            head := 0;
        END_IF;
        count := count - 1;
        status := 16#0000;
    END_IF;
END_IF;

elementCount := count;

(* ---- public-hard-04.candidate_02.st ---- *)
FUNCTION_BLOCK FB
VAR_INPUT
    enqueue : BOOL;
    dequeue : BOOL;
    reset : BOOL;
END_VAR
VAR_OUTPUT
    elementCount : DINT;
    status : WORD;
END_VAR
VAR_IN_OUT
    item : VARIANT;
    buffer : VARIANT;
END_VAR
VAR
    head : DINT := 0;
    tail : DINT := 0;
    count : DINT := 0;
    capacity : DINT := 0;
    elemSize : DINT := 0;
    initialized : BOOL := FALSE;
    prevEnqueue : BOOL := FALSE;
    prevDequeue : BOOL := FALSE;
    enqEdge : BOOL;
    deqEdge : BOOL;
    bufferAddr : PVOID;
    itemAddr : PVOID;
    bufferSize : DINT;
    itemSize : DINT;
    destAddr : PVOID;
    srcAddr : PVOID;
    copyLen : UDINT;
END_VAR

status := 16#0000;

IF NOT initialized THEN
    bufferSize := __VARINFO(buffer).diSize;
    itemSize := __VARINFO(item).diSize;
    IF (bufferSize > 0) AND (itemSize > 0) THEN
        elemSize := itemSize;
        capacity := bufferSize / elemSize;
        bufferAddr := __VARINFO(buffer).pvAddress;
        itemAddr := __VARINFO(item).pvAddress;
        head := 0;
        tail := 0;
        count := 0;
        initialized := TRUE;
    ELSE
        elementCount := 0;
        RETURN;
    END_IF;
END_IF;

enqEdge := enqueue AND NOT prevEnqueue;
deqEdge := dequeue AND NOT prevDequeue;
prevEnqueue := enqueue;
prevDequeue := dequeue;

IF reset THEN
    head := 0;
    tail := 0;
    count := 0;
    elementCount := 0;
    status := 16#0000;
    RETURN;
END_IF;

IF enqEdge THEN
    IF count >= capacity THEN
        status := 16#8002;
    ELSE
        destAddr := bufferAddr + (tail * elemSize);
        srcAddr := itemAddr;
        copyLen := TO_UDINT(elemSize);
        SysMemCpy(destAddr, srcAddr, copyLen);
        tail := tail + 1;
        IF tail >= capacity THEN
            tail := 0;
        END_IF;
        count := count + 1;
        status := 16#0000;
    END_IF;
END_IF;

IF deqEdge THEN
    IF count = 0 THEN
        status := 16#8001;
    ELSE
        srcAddr := bufferAddr + (head * elemSize);
        destAddr := itemAddr;
        copyLen := TO_UDINT(elemSize);
        SysMemCpy(destAddr, srcAddr, copyLen);
        head := head + 1;
        IF head >= capacity THEN
            head := 0;
        END_IF;
        count := count - 1;
        status := 16#0000;
    END_IF;
END_IF;

elementCount := count;

END_FUNCTION_BLOCK

(* ---- public-hard-04.raw_candidate_01.st ---- *)
FUNCTION_BLOCK FB
VAR_INPUT
    enqueue : BOOL;
    dequeue : BOOL;
    reset : BOOL;
END_VAR
VAR_OUTPUT
    elementCount : DINT;
    status : WORD;
END_VAR
VAR_IN_OUT
    item : VARIANT;
    buffer : VARIANT;
END_VAR
VAR
    head : DINT := 0;
    tail : DINT := 0;
    count : DINT := 0;
    capacity : DINT := 0;
    elemSize : DINT := 0;
    initialized : BOOL := FALSE;
    prevEnqueue : BOOL := FALSE;
    prevDequeue : BOOL := FALSE;
    enqEdge : BOOL;
    deqEdge : BOOL;
    bufferAddr : PVOID;
    itemAddr : PVOID;
    bufferSize : DINT;
    itemSize : DINT;
    destAddr : PVOID;
    srcAddr : PVOID;
    copyLen : UDINT;
END_VAR

status := 16#0000;

IF NOT initialized THEN
    bufferSize := __VARINFO(buffer).diSize;
    itemSize := __VARINFO(item).diSize;
    IF (bufferSize > 0) AND (itemSize > 0) THEN
        elemSize := itemSize;
        capacity := bufferSize / elemSize;
        bufferAddr := __VARINFO(buffer).pvAddress;
        itemAddr := __VARINFO(item).pvAddress;
        head := 0;
        tail := 0;
        count := 0;
        initialized := TRUE;
    ELSE
        elementCount := 0;
        RETURN;
    END_IF;
END_IF;

enqEdge := enqueue AND NOT prevEnqueue;
deqEdge := dequeue AND NOT prevDequeue;
prevEnqueue := enqueue;
prevDequeue := dequeue;

IF reset THEN
    head := 0;
    tail := 0;
    count := 0;
    elementCount := 0;
    status := 16#0000;
    RETURN;
END_IF;

IF enqEdge THEN
    IF count >= capacity THEN
        status := 16#8002;
    ELSE
        destAddr := bufferAddr + (tail * elemSize);
        srcAddr := itemAddr;
        copyLen := TO_UDINT(elemSize);
        SysMemCpy(destAddr, srcAddr, copyLen);
        tail := tail + 1;
        IF tail >= capacity THEN
            tail := 0;
        END_IF;
        count := count + 1;
        status := 16#0000;
    END_IF;
END_IF;

IF deqEdge THEN
    IF count = 0 THEN
        status := 16#8001;
    ELSE
        srcAddr := bufferAddr + (head * elemSize);
        destAddr := itemAddr;
        copyLen := TO_UDINT(elemSize);
        SysMemCpy(destAddr, srcAddr, copyLen);
        head := head + 1;
        IF head >= capacity THEN
            head := 0;
        END_IF;
        count := count - 1;
        status := 16#0000;
    END_IF;
END_IF;

elementCount := count;

(* ---- public-hard-04.raw_candidate_02.st ---- *)
FUNCTION_BLOCK FB
VAR_INPUT
    enqueue : BOOL;
    dequeue : BOOL;
    reset : BOOL;
END_VAR
VAR_OUTPUT
    elementCount : DINT;
    status : WORD;
END_VAR
VAR_IN_OUT
    item : VARIANT;
    buffer : VARIANT;
END_VAR
VAR
    head : DINT := 0;
    tail : DINT := 0;
    count : DINT := 0;
    capacity : DINT := 0;
    elemSize : DINT := 0;
    initialized : BOOL := FALSE;
    prevEnqueue : BOOL := FALSE;
    prevDequeue : BOOL := FALSE;
    enqEdge : BOOL;
    deqEdge : BOOL;
    bufferAddr : PVOID;
    itemAddr : PVOID;
    bufferSize : DINT;
    itemSize : DINT;
    destAddr : PVOID;
    srcAddr : PVOID;
    copyLen : UDINT;
END_VAR

status := 16#0000;

IF NOT initialized THEN
    bufferSize := __VARINFO(buffer).diSize;
    itemSize := __VARINFO(item).diSize;
    IF (bufferSize > 0) AND (itemSize > 0) THEN
        elemSize := itemSize;
        capacity := bufferSize / elemSize;
        bufferAddr := __VARINFO(buffer).pvAddress;
        itemAddr := __VARINFO(item).pvAddress;
        head := 0;
        tail := 0;
        count := 0;
        initialized := TRUE;
    ELSE
        elementCount := 0;
        RETURN;
    END_IF;
END_IF;

enqEdge := enqueue AND NOT prevEnqueue;
deqEdge := dequeue AND NOT prevDequeue;
prevEnqueue := enqueue;
prevDequeue := dequeue;

IF reset THEN
    head := 0;
    tail := 0;
    count := 0;
    elementCount := 0;
    status := 16#0000;
    RETURN;
END_IF;

IF enqEdge THEN
    IF count >= capacity THEN
        status := 16#8002;
    ELSE
        destAddr := bufferAddr + (tail * elemSize);
        srcAddr := itemAddr;
        copyLen := TO_UDINT(elemSize);
        SysMemCpy(destAddr, srcAddr, copyLen);
        tail := tail + 1;
        IF tail >= capacity THEN
            tail := 0;
        END_IF;
        count := count + 1;
        status := 16#0000;
    END_IF;
END_IF;

IF deqEdge THEN
    IF count = 0 THEN
        status := 16#8001;
    ELSE
        srcAddr := bufferAddr + (head * elemSize);
        destAddr := itemAddr;
        copyLen := TO_UDINT(elemSize);
        SysMemCpy(destAddr, srcAddr, copyLen);
        head := head + 1;
        IF head >= capacity THEN
            head := 0;
        END_IF;
        count := count - 1;
        status := 16#0000;
    END_IF;
END_IF;

elementCount := count;

END_FUNCTION_BLOCK

(* ---- public-hard-05.candidate_01.st ---- *)
FUNCTION_BLOCK MechanicalArmControl
VAR
    Step: INT := 1;                     // Current action step (1..8)
    ActionActive: BOOL := FALSE;        // TRUE when an automated action is being executed
    WaitingForStart: BOOL := TRUE;      // TRUE in single-step mode when waiting for start press
    CycleRunning: BOOL := FALSE;        // TRUE when a cycle is in progress (single/continuous)
    StartPrev: BOOL := FALSE;           // Previous value of Start input for edge detection
    StartPulse: BOOL := FALSE;          // One-scan pulse on rising edge of Start
    WaitingForStartPrev: BOOL := TRUE;  // Snapshot of WaitingForStart at scan start
    CycleRunningPrev: BOOL := FALSE;    // Snapshot of CycleRunning at scan start
END_VAR

// Rising edge detection for Start
StartPulse := Start AND NOT StartPrev;
StartPrev := Start;

// Capture previous states before any logic changes (to avoid race conditions)
WaitingForStartPrev := WaitingForStart;
CycleRunningPrev := CycleRunning;

IF NOT EmergencyStop THEN
    // Emergency stop triggered: stop all actions and reset automated state
    MoveDown := FALSE;
    MoveUp := FALSE;
    MoveLeft := FALSE;
    MoveRight := FALSE;
    ActivateGrip := FALSE;
    ActivateRelease := FALSE;
    Step := 1;
    ActionActive := FALSE;
    WaitingForStart := TRUE;
    CycleRunning := FALSE;
ELSE
    // Normal operation (no emergency stop)
    IF ManualMode THEN
        // Manual mode: direct button control with limit switch interlock
        MoveDown := DownButton AND NOT DownLimitSwitch;
        MoveUp := UpButton AND NOT UpLimitSwitch;
        MoveLeft := LeftButton AND NOT LeftLimitSwitch;
        MoveRight := RightButton AND NOT RightLimitSwitch;
        ActivateGrip := GripButton AND NOT GripLimitSwitch;
        ActivateRelease := ReleaseButton AND NOT ReleaseLimitSwitch;
        // Reset automated state when in manual mode
        Step := 1;
        ActionActive := FALSE;
        WaitingForStart := TRUE;
        CycleRunning := FALSE;
    ELSIF SingleStepMode THEN
        // Single step mode: one action per start press
        // Default outputs to false
        MoveDown := FALSE;
        MoveUp := FALSE;
        MoveLeft := FALSE;
        MoveRight := FALSE;
        ActivateGrip := FALSE;
        ActivateRelease := FALSE;

        // Start next action if waiting and start pulse occurs
        IF WaitingForStartPrev AND StartPulse THEN
            WaitingForStart := FALSE;
            ActionActive := TRUE;
            Step := 1;  // Always start from step 1
        END_IF;

        // Check completion of current action
        IF ActionActive THEN
            CASE Step OF
                1: IF DownLimitSwitch THEN
                       ActionActive := FALSE;
                       WaitingForStart := TRUE;
                       Step := 1;
                   END_IF;
                2: IF GripLimitSwitch THEN
                       ActionActive := FALSE;
                       WaitingForStart := TRUE;
                       Step := 2;
                   END_IF;
                3: IF UpLimitSwitch THEN
                       ActionActive := FALSE;
                       WaitingForStart := TRUE;
                       Step := 3;
                   END_IF;
                4: IF RightLimitSwitch THEN
                       ActionActive := FALSE;
                       WaitingForStart := TRUE;
                       Step := 4;
                   END_IF;
                5: IF DownLimitSwitch THEN
                       ActionActive := FALSE;
                       WaitingForStart := TRUE;
                       Step := 5;
                   END_IF;
                6: IF ReleaseLimitSwitch THEN
                       ActionActive := FALSE;
                       WaitingForStart := TRUE;
                       Step := 6;
                   END_IF;
                7: IF UpLimitSwitch THEN
                       ActionActive := FALSE;
                       WaitingForStart := TRUE;
                       Step := 7;
                   END_IF;
                8: IF LeftLimitSwitch THEN
                       ActionActive := FALSE;
                       WaitingForStart := TRUE;
                       Step := 1;  // Reset to step 1 for next cycle
                   END_IF;
            END_CASE;
        END_IF;

        // Set outputs based on current step and action active
        IF ActionActive THEN
            CASE Step OF
                1: MoveDown := TRUE;
                2: ActivateGrip := TRUE;
                3: MoveUp := TRUE;
                4: MoveRight := TRUE;
                5: MoveDown := TRUE;
                6: ActivateRelease := TRUE;
                7: MoveUp := TRUE;
                8: MoveLeft := TRUE;
            END_CASE;
        END_IF;
    ELSIF SingleCycleMode THEN
        // Single cycle mode: complete one full cycle automatically
        MoveDown := FALSE;
        MoveUp := FALSE;
        MoveLeft := FALSE;
        MoveRight := FALSE;
        ActivateGrip := FALSE;
        ActivateRelease := FALSE;

        // Start cycle on rising edge of Start if not already running
        IF NOT CycleRunningPrev AND StartPulse THEN
            CycleRunning := TRUE;
            Step := 1;
            ActionActive := TRUE;
        END_IF;

        // Execute cycle and advance to next action on completion
        IF CycleRunning AND ActionActive THEN
            CASE Step OF
                1: IF DownLimitSwitch THEN Step := 2; END_IF;
                2: IF GripLimitSwitch THEN Step := 3; END_IF;
                3: IF UpLimitSwitch THEN Step := 4; END_IF;
                4: IF RightLimitSwitch THEN Step := 5; END_IF;
                5: IF DownLimitSwitch THEN Step := 6; END_IF;
                6: IF ReleaseLimitSwitch THEN Step := 7; END_IF;
                7: IF UpLimitSwitch THEN Step := 8; END_IF;
                8: IF LeftLimitSwitch THEN
                       ActionActive := FALSE;   // Cycle finished
                       CycleRunning := FALSE;
                       Step := 1;               // Reset for next start
                   END_IF;
            END_CASE;
        END_IF;

        // Set outputs according to current step
        IF CycleRunning AND ActionActive THEN
            CASE Step OF
                1: MoveDown := TRUE;
                2: ActivateGrip := TRUE;
                3: MoveUp := TRUE;
                4: MoveRight := TRUE;
                5: MoveDown := TRUE;
                6: ActivateRelease := TRUE;
                7: MoveUp := TRUE;
                8: MoveLeft := TRUE;
            END_CASE;
        END_IF;
    ELSIF ContinuousMode THEN
        // Continuous mode: repeat cycle indefinitely
        MoveDown := FALSE;
        MoveUp := FALSE;
        MoveLeft := FALSE;
        MoveRight := FALSE;
        ActivateGrip := FALSE;
        ActivateRelease := FALSE;

        // Start continuous operation on rising edge of Start if not already running
        IF NOT CycleRunningPrev AND StartPulse THEN
            CycleRunning := TRUE;
            Step := 1;
            ActionActive := TRUE;
        END_IF;

        // Execute cycle and loop back to step 1 after step 8
        IF CycleRunning AND ActionActive THEN
            CASE Step OF
                1: IF DownLimitSwitch THEN Step := 2; END_IF;
                2: IF GripLimitSwitch THEN Step := 3; END_IF;
                3: IF UpLimitSwitch THEN Step := 4; END_IF;
                4: IF RightLimitSwitch THEN Step := 5; END_IF;
                5: IF DownLimitSwitch THEN Step := 6; END_IF;
                6: IF ReleaseLimitSwitch THEN Step := 7; END_IF;
                7: IF UpLimitSwitch THEN Step := 8; END_IF;
                8: IF LeftLimitSwitch THEN Step := 1; END_IF;  // Loop back
            END_CASE;
        END_IF;

        // Set outputs according to current step
        IF CycleRunning AND ActionActive THEN
            CASE Step OF
                1: MoveDown := TRUE;
                2: ActivateGrip := TRUE;
                3: MoveUp := TRUE;
                4: MoveRight := TRUE;
                5: MoveDown := TRUE;
                6: ActivateRelease := TRUE;
                7: MoveUp := TRUE;
                8: MoveLeft := TRUE;
            END_CASE;
        END_IF;
    ELSE
        // No mode selected (should not happen, but safe default)
        MoveDown := FALSE;
        MoveUp := FALSE;
        MoveLeft := FALSE;
        MoveRight := FALSE;
        ActivateGrip := FALSE;
        ActivateRelease := FALSE;
        Step := 1;
        ActionActive := FALSE;
        WaitingForStart := TRUE;
        CycleRunning := FALSE;
    END_IF;
END_IF;

(* ---- public-hard-05.candidate_02.st ---- *)
FUNCTION_BLOCK MechanicalArmControl
VAR
    Step: INT := 1;                     // Current action step (1..8)
    ActionActive: BOOL := FALSE;        // TRUE when an automated action is being executed
    WaitingForStart: BOOL := TRUE;      // TRUE in single-step mode when waiting for start press
    CycleRunning: BOOL := FALSE;        // TRUE when a cycle is in progress (single/continuous)
    StartPrev: BOOL := FALSE;           // Previous value of Start input for edge detection
    StartPulse: BOOL := FALSE;          // One-scan pulse on rising edge of Start
    WaitingForStartPrev: BOOL := TRUE;  // Snapshot of WaitingForStart at scan start
    CycleRunningPrev: BOOL := FALSE;    // Snapshot of CycleRunning at scan start
END_VAR

// Rising edge detection for Start
StartPulse := Start AND NOT StartPrev;
StartPrev := Start;

// Capture previous states before any logic changes (to avoid race conditions)
WaitingForStartPrev := WaitingForStart;
CycleRunningPrev := CycleRunning;

IF NOT EmergencyStop THEN
    // Emergency stop triggered: stop all actions and reset automated state
    MoveDown := FALSE;
    MoveUp := FALSE;
    MoveLeft := FALSE;
    MoveRight := FALSE;
    ActivateGrip := FALSE;
    ActivateRelease := FALSE;
    Step := 1;
    ActionActive := FALSE;
    WaitingForStart := TRUE;
    CycleRunning := FALSE;
ELSE
    // Normal operation (no emergency stop)
    IF ManualMode THEN
        // Manual mode: direct button control with limit switch interlock
        MoveDown := DownButton AND NOT DownLimitSwitch;
        MoveUp := UpButton AND NOT UpLimitSwitch;
        MoveLeft := LeftButton AND NOT LeftLimitSwitch;
        MoveRight := RightButton AND NOT RightLimitSwitch;
        ActivateGrip := GripButton AND NOT GripLimitSwitch;
        ActivateRelease := ReleaseButton AND NOT ReleaseLimitSwitch;
        // Reset automated state when in manual mode
        Step := 1;
        ActionActive := FALSE;
        WaitingForStart := TRUE;
        CycleRunning := FALSE;
    ELSIF SingleStepMode THEN
        // Single step mode: one action per start press
        MoveDown := FALSE;
        MoveUp := FALSE;
        MoveLeft := FALSE;
        MoveRight := FALSE;
        ActivateGrip := FALSE;
        ActivateRelease := FALSE;

        IF WaitingForStartPrev AND StartPulse THEN
            WaitingForStart := FALSE;
            ActionActive := TRUE;
            Step := 1;  // Always start from step 1
        END_IF;

        IF ActionActive THEN
            CASE Step OF
                1: IF DownLimitSwitch THEN
                       ActionActive := FALSE;
                       WaitingForStart := TRUE;
                       Step := 1;
                   END_IF;
                2: IF GripLimitSwitch THEN
                       ActionActive := FALSE;
                       WaitingForStart := TRUE;
                       Step := 2;
                   END_IF;
                3: IF UpLimitSwitch THEN
                       ActionActive := FALSE;
                       WaitingForStart := TRUE;
                       Step := 3;
                   END_IF;
                4: IF RightLimitSwitch THEN
                       ActionActive := FALSE;
                       WaitingForStart := TRUE;
                       Step := 4;
                   END_IF;
                5: IF DownLimitSwitch THEN
                       ActionActive := FALSE;
                       WaitingForStart := TRUE;
                       Step := 5;
                   END_IF;
                6: IF ReleaseLimitSwitch THEN
                       ActionActive := FALSE;
                       WaitingForStart := TRUE;
                       Step := 6;
                   END_IF;
                7: IF UpLimitSwitch THEN
                       ActionActive := FALSE;
                       WaitingForStart := TRUE;
                       Step := 7;
                   END_IF;
                8: IF LeftLimitSwitch THEN
                       ActionActive := FALSE;
                       WaitingForStart := TRUE;
                       Step := 1;  // Reset to step 1 for next cycle
                   END_IF;
            END_CASE;
        END_IF;

        IF ActionActive THEN
            CASE Step OF
                1: MoveDown := TRUE;
                2: ActivateGrip := TRUE;
                3: MoveUp := TRUE;
                4: MoveRight := TRUE;
                5: MoveDown := TRUE;
                6: ActivateRelease := TRUE;
                7: MoveUp := TRUE;
                8: MoveLeft := TRUE;
            END_CASE;
        END_IF;
    ELSIF SingleCycleMode THEN
        // Single cycle mode: complete one full cycle automatically
        MoveDown := FALSE;
        MoveUp := FALSE;
        MoveLeft := FALSE;
        MoveRight := FALSE;
        ActivateGrip := FALSE;
        ActivateRelease := FALSE;

        IF NOT CycleRunningPrev AND StartPulse THEN
            CycleRunning := TRUE;
            Step := 1;
            ActionActive := TRUE;
        END_IF;

        IF CycleRunning AND ActionActive THEN
            CASE Step OF
                1: IF DownLimitSwitch THEN Step := 2; END_IF;
                2: IF GripLimitSwitch THEN Step := 3; END_IF;
                3: IF UpLimitSwitch THEN Step := 4; END_IF;
                4: IF RightLimitSwitch THEN Step := 5; END_IF;
                5: IF DownLimitSwitch THEN Step := 6; END_IF;
                6: IF ReleaseLimitSwitch THEN Step := 7; END_IF;
                7: IF UpLimitSwitch THEN Step := 8; END_IF;
                8: IF LeftLimitSwitch THEN
                       ActionActive := FALSE;   // Cycle finished
                       CycleRunning := FALSE;
                       Step := 1;               // Reset for next start
                   END_IF;
            END_CASE;
        END_IF;

        IF CycleRunning AND ActionActive THEN
            CASE Step OF
                1: MoveDown := TRUE;
                2: ActivateGrip := TRUE;
                3: MoveUp := TRUE;
                4: MoveRight := TRUE;
                5: MoveDown := TRUE;
                6: ActivateRelease := TRUE;
                7: MoveUp := TRUE;
                8: MoveLeft := TRUE;
            END_CASE;
        END_IF;
    ELSIF ContinuousMode THEN
        // Continuous mode: repeat cycle indefinitely
        MoveDown := FALSE;
        MoveUp := FALSE;
        MoveLeft := FALSE;
        MoveRight := FALSE;
        ActivateGrip := FALSE;
        ActivateRelease := FALSE;

        IF NOT CycleRunningPrev AND StartPulse THEN
            CycleRunning := TRUE;
            Step := 1;
            ActionActive := TRUE;
        END_IF;

        IF CycleRunning AND ActionActive THEN
            CASE Step OF
                1: IF DownLimitSwitch THEN Step := 2; END_IF;
                2: IF GripLimitSwitch THEN Step := 3; END_IF;
                3: IF UpLimitSwitch THEN Step := 4; END_IF;
                4: IF RightLimitSwitch THEN Step := 5; END_IF;
                5: IF DownLimitSwitch THEN Step := 6; END_IF;
                6: IF ReleaseLimitSwitch THEN Step := 7; END_IF;
                7: IF UpLimitSwitch THEN Step := 8; END_IF;
                8: IF LeftLimitSwitch THEN Step := 1; END_IF;  // Loop back
            END_CASE;
        END_IF;

        IF CycleRunning AND ActionActive THEN
            CASE Step OF
                1: MoveDown := TRUE;
                2: ActivateGrip := TRUE;
                3: MoveUp := TRUE;
                4: MoveRight := TRUE;
                5: MoveDown := TRUE;
                6: ActivateRelease := TRUE;
                7: MoveUp := TRUE;
                8: MoveLeft := TRUE;
            END_CASE;
        END_IF;
    ELSE
        // No mode selected (should not happen, but safe default)
        MoveDown := FALSE;
        MoveUp := FALSE;
        MoveLeft := FALSE;
        MoveRight := FALSE;
        ActivateGrip := FALSE;
        ActivateRelease := FALSE;
        Step := 1;
        ActionActive := FALSE;
        WaitingForStart := TRUE;
        CycleRunning := FALSE;
    END_IF;
END_IF;

END_FUNCTION_BLOCK

(* ---- public-hard-05.raw_candidate_01.st ---- *)
FUNCTION_BLOCK MechanicalArmControl
VAR
    Step: INT := 1;                     // Current action step (1..8)
    ActionActive: BOOL := FALSE;        // TRUE when an automated action is being executed
    WaitingForStart: BOOL := TRUE;      // TRUE in single-step mode when waiting for start press
    CycleRunning: BOOL := FALSE;        // TRUE when a cycle is in progress (single/continuous)
    StartPrev: BOOL := FALSE;           // Previous value of Start input for edge detection
    StartPulse: BOOL := FALSE;          // One-scan pulse on rising edge of Start
    WaitingForStartPrev: BOOL := TRUE;  // Snapshot of WaitingForStart at scan start
    CycleRunningPrev: BOOL := FALSE;    // Snapshot of CycleRunning at scan start
END_VAR

// Rising edge detection for Start
StartPulse := Start AND NOT StartPrev;
StartPrev := Start;

// Capture previous states before any logic changes (to avoid race conditions)
WaitingForStartPrev := WaitingForStart;
CycleRunningPrev := CycleRunning;

IF NOT EmergencyStop THEN
    // Emergency stop triggered: stop all actions and reset automated state
    MoveDown := FALSE;
    MoveUp := FALSE;
    MoveLeft := FALSE;
    MoveRight := FALSE;
    ActivateGrip := FALSE;
    ActivateRelease := FALSE;
    Step := 1;
    ActionActive := FALSE;
    WaitingForStart := TRUE;
    CycleRunning := FALSE;
ELSE
    // Normal operation (no emergency stop)
    IF ManualMode THEN
        // Manual mode: direct button control with limit switch interlock
        MoveDown := DownButton AND NOT DownLimitSwitch;
        MoveUp := UpButton AND NOT UpLimitSwitch;
        MoveLeft := LeftButton AND NOT LeftLimitSwitch;
        MoveRight := RightButton AND NOT RightLimitSwitch;
        ActivateGrip := GripButton AND NOT GripLimitSwitch;
        ActivateRelease := ReleaseButton AND NOT ReleaseLimitSwitch;
        // Reset automated state when in manual mode
        Step := 1;
        ActionActive := FALSE;
        WaitingForStart := TRUE;
        CycleRunning := FALSE;
    ELSIF SingleStepMode THEN
        // Single step mode: one action per start press
        // Default outputs to false
        MoveDown := FALSE;
        MoveUp := FALSE;
        MoveLeft := FALSE;
        MoveRight := FALSE;
        ActivateGrip := FALSE;
        ActivateRelease := FALSE;

        // Start next action if waiting and start pulse occurs
        IF WaitingForStartPrev AND StartPulse THEN
            WaitingForStart := FALSE;
            ActionActive := TRUE;
            Step := 1;  // Always start from step 1
        END_IF;

        // Check completion of current action
        IF ActionActive THEN
            CASE Step OF
                1: IF DownLimitSwitch THEN
                       ActionActive := FALSE;
                       WaitingForStart := TRUE;
                       Step := 1;
                   END_IF;
                2: IF GripLimitSwitch THEN
                       ActionActive := FALSE;
                       WaitingForStart := TRUE;
                       Step := 2;
                   END_IF;
                3: IF UpLimitSwitch THEN
                       ActionActive := FALSE;
                       WaitingForStart := TRUE;
                       Step := 3;
                   END_IF;
                4: IF RightLimitSwitch THEN
                       ActionActive := FALSE;
                       WaitingForStart := TRUE;
                       Step := 4;
                   END_IF;
                5: IF DownLimitSwitch THEN
                       ActionActive := FALSE;
                       WaitingForStart := TRUE;
                       Step := 5;
                   END_IF;
                6: IF ReleaseLimitSwitch THEN
                       ActionActive := FALSE;
                       WaitingForStart := TRUE;
                       Step := 6;
                   END_IF;
                7: IF UpLimitSwitch THEN
                       ActionActive := FALSE;
                       WaitingForStart := TRUE;
                       Step := 7;
                   END_IF;
                8: IF LeftLimitSwitch THEN
                       ActionActive := FALSE;
                       WaitingForStart := TRUE;
                       Step := 1;  // Reset to step 1 for next cycle
                   END_IF;
            END_CASE;
        END_IF;

        // Set outputs based on current step and action active
        IF ActionActive THEN
            CASE Step OF
                1: MoveDown := TRUE;
                2: ActivateGrip := TRUE;
                3: MoveUp := TRUE;
                4: MoveRight := TRUE;
                5: MoveDown := TRUE;
                6: ActivateRelease := TRUE;
                7: MoveUp := TRUE;
                8: MoveLeft := TRUE;
            END_CASE;
        END_IF;
    ELSIF SingleCycleMode THEN
        // Single cycle mode: complete one full cycle automatically
        MoveDown := FALSE;
        MoveUp := FALSE;
        MoveLeft := FALSE;
        MoveRight := FALSE;
        ActivateGrip := FALSE;
        ActivateRelease := FALSE;

        // Start cycle on rising edge of Start if not already running
        IF NOT CycleRunningPrev AND StartPulse THEN
            CycleRunning := TRUE;
            Step := 1;
            ActionActive := TRUE;
        END_IF;

        // Execute cycle and advance to next action on completion
        IF CycleRunning AND ActionActive THEN
            CASE Step OF
                1: IF DownLimitSwitch THEN Step := 2; END_IF;
                2: IF GripLimitSwitch THEN Step := 3; END_IF;
                3: IF UpLimitSwitch THEN Step := 4; END_IF;
                4: IF RightLimitSwitch THEN Step := 5; END_IF;
                5: IF DownLimitSwitch THEN Step := 6; END_IF;
                6: IF ReleaseLimitSwitch THEN Step := 7; END_IF;
                7: IF UpLimitSwitch THEN Step := 8; END_IF;
                8: IF LeftLimitSwitch THEN
                       ActionActive := FALSE;   // Cycle finished
                       CycleRunning := FALSE;
                       Step := 1;               // Reset for next start
                   END_IF;
            END_CASE;
        END_IF;

        // Set outputs according to current step
        IF CycleRunning AND ActionActive THEN
            CASE Step OF
                1: MoveDown := TRUE;
                2: ActivateGrip := TRUE;
                3: MoveUp := TRUE;
                4: MoveRight := TRUE;
                5: MoveDown := TRUE;
                6: ActivateRelease := TRUE;
                7: MoveUp := TRUE;
                8: MoveLeft := TRUE;
            END_CASE;
        END_IF;
    ELSIF ContinuousMode THEN
        // Continuous mode: repeat cycle indefinitely
        MoveDown := FALSE;
        MoveUp := FALSE;
        MoveLeft := FALSE;
        MoveRight := FALSE;
        ActivateGrip := FALSE;
        ActivateRelease := FALSE;

        // Start continuous operation on rising edge of Start if not already running
        IF NOT CycleRunningPrev AND StartPulse THEN
            CycleRunning := TRUE;
            Step := 1;
            ActionActive := TRUE;
        END_IF;

        // Execute cycle and loop back to step 1 after step 8
        IF CycleRunning AND ActionActive THEN
            CASE Step OF
                1: IF DownLimitSwitch THEN Step := 2; END_IF;
                2: IF GripLimitSwitch THEN Step := 3; END_IF;
                3: IF UpLimitSwitch THEN Step := 4; END_IF;
                4: IF RightLimitSwitch THEN Step := 5; END_IF;
                5: IF DownLimitSwitch THEN Step := 6; END_IF;
                6: IF ReleaseLimitSwitch THEN Step := 7; END_IF;
                7: IF UpLimitSwitch THEN Step := 8; END_IF;
                8: IF LeftLimitSwitch THEN Step := 1; END_IF;  // Loop back
            END_CASE;
        END_IF;

        // Set outputs according to current step
        IF CycleRunning AND ActionActive THEN
            CASE Step OF
                1: MoveDown := TRUE;
                2: ActivateGrip := TRUE;
                3: MoveUp := TRUE;
                4: MoveRight := TRUE;
                5: MoveDown := TRUE;
                6: ActivateRelease := TRUE;
                7: MoveUp := TRUE;
                8: MoveLeft := TRUE;
            END_CASE;
        END_IF;
    ELSE
        // No mode selected (should not happen, but safe default)
        MoveDown := FALSE;
        MoveUp := FALSE;
        MoveLeft := FALSE;
        MoveRight := FALSE;
        ActivateGrip := FALSE;
        ActivateRelease := FALSE;
        Step := 1;
        ActionActive := FALSE;
        WaitingForStart := TRUE;
        CycleRunning := FALSE;
    END_IF;
END_IF;
